(* Logix 5000 project; controller CIP vendor 1 type 14 code 106 rev 20.12; software revision 20.06; part 2 of 13 *)
(* tags used below, declared in another part *)
   Bit : BOOL[128];
   Counter : COUNTER[10];
   IN_N7_100_199 : INT[100];
   Integer : DINT[150];
   Integer_1 : ALIAS FOR Integer[1];
   Level_Bits : BOOL[32];
   One_Shot : BOOL[128];
   OpCode_Pin : DINT[5];
   OpCode_Word : DINT[5,97];
   Panelview : INT[40];
   PV_Security : Security_Main_HMI;
   Recipe : RECIPE[41];

        [24].Setpoint[26] := 9.0, [24].Setpoint[27] := 10.0, [24].Setpoint[28] := 50.0, [24].Setpoint[29] := 3.0, [24].Setpoint[30] := 17.0, [24].Setpoint[31] := 300.0, [24].Setpoint[32] := 2.0, [24].Setpoint[33] := 2.0, [24].Setpoint[34] := 900.0, [24].Setpoint[37] := 70.0, [24].Setpoint[38] := 100.0, [24].Setpoint[39] := 110.0, [24].Setpoint[40] := 30.0, [24].Setpoint[41] := 60.0, [24].Setpoint[42] := 60.0, [24].Setpoint[43] := 3000.0, [24].Setpoint[44] := 300.0, [24].Setpoint[45] := 185.0, [24].Setpoint[46] := 10.0, [24].Setpoint[47] := 25.0, [24].Setpoint[48] := 150.0, [24].Setpoint[49] := 125.0, [24].Setpoint[50] := 100.0, [24].Setpoint[51] := 80.0, [24].Setpoint[52] := 100.0, [24].Setpoint[53] := 50.0, [24].Setpoint[54] := 85.0, [24].Setpoint[55] := 40.0, [24].Setpoint[56] := 60.0, [24].Setpoint[57] := 90.0, [24].Setpoint[58] := 4.0, [24].Setpoint[61] := 10.0, [24].Setpoint[62] := 1.0, [24].Setpoint[65] := 100.0, [24].Setpoint[66] := 15.0, [24].Setpoint[67] := 50.0, [24].Setpoint[68] := 5.0, [24].Setpoint[69] := 100.0, [24].Setpoint[70] := 15.0, [24].Setpoint[71] := 100.0, [24].Setpoint[72] := 15.0, [24].Setpoint[73] := 120.0, [24].Setpoint[74] := 20.0, [24].Setpoint[75] := 120.0, [24].Setpoint[76] := 20.0, [24].Setpoint[77] := 100.0, [24].Setpoint[78] := 15.0, [24].Setpoint[79] := 100.0, [24].Setpoint[80] := 15.0, [24].Setpoint[81] := 45.0, [24].Setpoint[82] := 30.0, [24].Setpoint[83] := 5.0, [24].Setpoint[85] := 5.0, [24].Setpoint[86] := 9.0, [24].Setpoint[92] := 75.0, [24].Setpoint[93] := 90.0, [24].Setpoint[94] := 5.0, [24].Setpoint[95] := 110.0, [24].Setpoint[96] := 10.0, [24].Name := 'RECIPE #24',
        [25].Setpoint[1] := 55.0, [25].Setpoint[2] := 65.0, [25].Setpoint[3] := 60.0, [25].Setpoint[4] := 45.0, [25].Setpoint[5] := 65.0, [25].Setpoint[6] := 25.0, [25].Setpoint[7] := 53.0, [25].Setpoint[8] := 63.0, [25].Setpoint[9] := 57.0, [25].Setpoint[10] := 43.0, [25].Setpoint[11] := 63.0, [25].Setpoint[12] := 22.0, [25].Setpoint[13] := 85.0, [25].Setpoint[14] := 900.0, [25].Setpoint[15] := 300.0, [25].Setpoint[16] := 300.0, [25].Setpoint[17] := 15.0, [25].Setpoint[18] := 14.0, [25].Setpoint[19] := 15.0, [25].Setpoint[20] := 45.0, [25].Setpoint[21] := 5.0, [25].Setpoint[22] := 15.0, [25].Setpoint[23] := 300.0, [25].Setpoint[24] := 2.0, [25].Setpoint[25] := 10.0, [25].Setpoint[26] := 9.0, [25].Setpoint[27] := 10.0, [25].Setpoint[28] := 50.0, [25].Setpoint[29] := 3.0, [25].Setpoint[30] := 17.0, [25].Setpoint[31] := 300.0, [25].Setpoint[32] := 2.0, [25].Setpoint[33] := 2.0, [25].Setpoint[34] := 900.0, [25].Setpoint[37] := 70.0, [25].Setpoint[38] := 100.0, [25].Setpoint[39] := 110.0, [25].Setpoint[40] := 30.0, [25].Setpoint[41] := 60.0, [25].Setpoint[42] := 60.0, [25].Setpoint[43] := 3000.0, [25].Setpoint[44] := 300.0, [25].Setpoint[45] := 185.0, [25].Setpoint[46] := 10.0, [25].Setpoint[47] := 25.0, [25].Setpoint[48] := 150.0, [25].Setpoint[49] := 125.0, [25].Setpoint[50] := 100.0, [25].Setpoint[51] := 80.0, [25].Setpoint[52] := 100.0, [25].Setpoint[53] := 50.0, [25].Setpoint[54] := 85.0, [25].Setpoint[55] := 40.0, [25].Setpoint[56] := 60.0, [25].Setpoint[57] := 90.0, [25].Setpoint[58] := 4.0, [25].Setpoint[61] := 10.0, [25].Setpoint[62] := 1.0, [25].Setpoint[65] := 100.0, [25].Setpoint[66] := 15.0,
        [25].Setpoint[67] := 50.0, [25].Setpoint[68] := 5.0, [25].Setpoint[69] := 100.0, [25].Setpoint[70] := 15.0, [25].Setpoint[71] := 100.0, [25].Setpoint[72] := 15.0, [25].Setpoint[73] := 120.0, [25].Setpoint[74] := 20.0, [25].Setpoint[75] := 120.0, [25].Setpoint[76] := 20.0, [25].Setpoint[77] := 100.0, [25].Setpoint[78] := 15.0, [25].Setpoint[79] := 100.0, [25].Setpoint[80] := 15.0, [25].Setpoint[81] := 45.0, [25].Setpoint[82] := 30.0, [25].Setpoint[83] := 5.0, [25].Setpoint[85] := 5.0, [25].Setpoint[86] := 9.0, [25].Setpoint[92] := 75.0, [25].Setpoint[93] := 90.0, [25].Setpoint[94] := 5.0, [25].Setpoint[95] := 110.0, [25].Setpoint[96] := 10.0, [25].Name := 'RECIPE #25', [26].Setpoint[1] := 55.0, [26].Setpoint[2] := 65.0, [26].Setpoint[3] := 60.0, [26].Setpoint[4] := 45.0, [26].Setpoint[5] := 65.0, [26].Setpoint[6] := 25.0, [26].Setpoint[7] := 53.0, [26].Setpoint[8] := 63.0, [26].Setpoint[9] := 57.0, [26].Setpoint[10] := 43.0, [26].Setpoint[11] := 63.0, [26].Setpoint[12] := 22.0, [26].Setpoint[13] := 85.0, [26].Setpoint[14] := 900.0, [26].Setpoint[15] := 300.0, [26].Setpoint[16] := 300.0, [26].Setpoint[17] := 15.0, [26].Setpoint[18] := 14.0, [26].Setpoint[19] := 15.0, [26].Setpoint[20] := 45.0, [26].Setpoint[21] := 5.0, [26].Setpoint[22] := 15.0, [26].Setpoint[23] := 300.0, [26].Setpoint[24] := 2.0, [26].Setpoint[25] := 10.0, [26].Setpoint[26] := 9.0, [26].Setpoint[27] := 10.0, [26].Setpoint[28] := 50.0, [26].Setpoint[29] := 3.0, [26].Setpoint[30] := 17.0, [26].Setpoint[31] := 300.0, [26].Setpoint[32] := 2.0, [26].Setpoint[33] := 2.0, [26].Setpoint[34] := 900.0, [26].Setpoint[37] := 70.0,
        [26].Setpoint[38] := 100.0, [26].Setpoint[39] := 110.0, [26].Setpoint[40] := 30.0, [26].Setpoint[41] := 60.0, [26].Setpoint[42] := 60.0, [26].Setpoint[43] := 3000.0, [26].Setpoint[44] := 300.0, [26].Setpoint[45] := 185.0, [26].Setpoint[46] := 10.0, [26].Setpoint[47] := 25.0, [26].Setpoint[48] := 150.0, [26].Setpoint[49] := 125.0, [26].Setpoint[50] := 100.0, [26].Setpoint[51] := 80.0, [26].Setpoint[52] := 100.0, [26].Setpoint[53] := 50.0, [26].Setpoint[54] := 85.0, [26].Setpoint[55] := 40.0, [26].Setpoint[56] := 60.0, [26].Setpoint[57] := 90.0, [26].Setpoint[58] := 4.0, [26].Setpoint[61] := 10.0, [26].Setpoint[62] := 1.0, [26].Setpoint[65] := 100.0, [26].Setpoint[66] := 15.0, [26].Setpoint[67] := 50.0, [26].Setpoint[68] := 5.0, [26].Setpoint[69] := 100.0, [26].Setpoint[70] := 15.0, [26].Setpoint[71] := 100.0, [26].Setpoint[72] := 15.0, [26].Setpoint[73] := 120.0, [26].Setpoint[74] := 20.0, [26].Setpoint[75] := 120.0, [26].Setpoint[76] := 20.0, [26].Setpoint[77] := 100.0, [26].Setpoint[78] := 15.0, [26].Setpoint[79] := 100.0, [26].Setpoint[80] := 15.0, [26].Setpoint[81] := 45.0, [26].Setpoint[82] := 30.0, [26].Setpoint[83] := 5.0, [26].Setpoint[85] := 5.0, [26].Setpoint[86] := 9.0, [26].Setpoint[92] := 75.0, [26].Setpoint[93] := 90.0, [26].Setpoint[94] := 5.0, [26].Setpoint[95] := 110.0, [26].Setpoint[96] := 10.0, [26].Name := 'RECIPE #26', [27].Setpoint[1] := 55.0, [27].Setpoint[2] := 65.0, [27].Setpoint[3] := 60.0, [27].Setpoint[4] := 45.0, [27].Setpoint[5] := 65.0, [27].Setpoint[6] := 25.0, [27].Setpoint[7] := 53.0, [27].Setpoint[8] := 63.0, [27].Setpoint[9] := 57.0, [27].Setpoint[10] := 43.0,
        [27].Setpoint[11] := 63.0, [27].Setpoint[12] := 22.0, [27].Setpoint[13] := 85.0, [27].Setpoint[14] := 900.0, [27].Setpoint[15] := 300.0, [27].Setpoint[16] := 300.0, [27].Setpoint[17] := 15.0, [27].Setpoint[18] := 14.0, [27].Setpoint[19] := 15.0, [27].Setpoint[20] := 45.0, [27].Setpoint[21] := 5.0, [27].Setpoint[22] := 15.0, [27].Setpoint[23] := 300.0, [27].Setpoint[24] := 2.0, [27].Setpoint[25] := 10.0, [27].Setpoint[26] := 9.0, [27].Setpoint[27] := 10.0, [27].Setpoint[28] := 50.0, [27].Setpoint[29] := 3.0, [27].Setpoint[30] := 17.0, [27].Setpoint[31] := 300.0, [27].Setpoint[32] := 2.0, [27].Setpoint[33] := 2.0, [27].Setpoint[34] := 900.0, [27].Setpoint[37] := 70.0, [27].Setpoint[38] := 100.0, [27].Setpoint[39] := 110.0, [27].Setpoint[40] := 30.0, [27].Setpoint[41] := 60.0, [27].Setpoint[42] := 60.0, [27].Setpoint[43] := 3000.0, [27].Setpoint[44] := 300.0, [27].Setpoint[45] := 185.0, [27].Setpoint[46] := 10.0, [27].Setpoint[47] := 25.0, [27].Setpoint[48] := 150.0, [27].Setpoint[49] := 125.0, [27].Setpoint[50] := 100.0, [27].Setpoint[51] := 80.0, [27].Setpoint[52] := 100.0, [27].Setpoint[53] := 50.0, [27].Setpoint[54] := 85.0, [27].Setpoint[55] := 40.0, [27].Setpoint[56] := 60.0, [27].Setpoint[57] := 90.0, [27].Setpoint[58] := 4.0, [27].Setpoint[61] := 10.0, [27].Setpoint[62] := 1.0, [27].Setpoint[65] := 100.0, [27].Setpoint[66] := 15.0, [27].Setpoint[67] := 50.0, [27].Setpoint[68] := 5.0, [27].Setpoint[69] := 100.0, [27].Setpoint[70] := 15.0, [27].Setpoint[71] := 100.0, [27].Setpoint[72] := 15.0, [27].Setpoint[73] := 120.0, [27].Setpoint[74] := 20.0, [27].Setpoint[75] := 120.0, [27].Setpoint[76] := 20.0,
        [27].Setpoint[77] := 100.0, [27].Setpoint[78] := 15.0, [27].Setpoint[79] := 100.0, [27].Setpoint[80] := 15.0, [27].Setpoint[81] := 45.0, [27].Setpoint[82] := 30.0, [27].Setpoint[83] := 5.0, [27].Setpoint[85] := 5.0, [27].Setpoint[86] := 9.0, [27].Setpoint[92] := 75.0, [27].Setpoint[93] := 90.0, [27].Setpoint[94] := 5.0, [27].Setpoint[95] := 110.0, [27].Setpoint[96] := 10.0, [27].Name := 'RECIPE #27', [28].Setpoint[1] := 55.0, [28].Setpoint[2] := 65.0, [28].Setpoint[3] := 60.0, [28].Setpoint[4] := 45.0, [28].Setpoint[5] := 65.0, [28].Setpoint[6] := 25.0, [28].Setpoint[7] := 53.0, [28].Setpoint[8] := 63.0, [28].Setpoint[9] := 57.0, [28].Setpoint[10] := 43.0, [28].Setpoint[11] := 63.0, [28].Setpoint[12] := 22.0, [28].Setpoint[13] := 85.0, [28].Setpoint[14] := 900.0, [28].Setpoint[15] := 300.0, [28].Setpoint[16] := 300.0, [28].Setpoint[17] := 15.0, [28].Setpoint[18] := 14.0, [28].Setpoint[19] := 15.0, [28].Setpoint[20] := 45.0, [28].Setpoint[21] := 5.0, [28].Setpoint[22] := 15.0, [28].Setpoint[23] := 300.0, [28].Setpoint[24] := 2.0, [28].Setpoint[25] := 10.0, [28].Setpoint[26] := 9.0, [28].Setpoint[27] := 10.0, [28].Setpoint[28] := 50.0, [28].Setpoint[29] := 3.0, [28].Setpoint[30] := 17.0, [28].Setpoint[31] := 300.0, [28].Setpoint[32] := 2.0, [28].Setpoint[33] := 2.0, [28].Setpoint[34] := 900.0, [28].Setpoint[37] := 70.0, [28].Setpoint[38] := 100.0, [28].Setpoint[39] := 110.0, [28].Setpoint[40] := 30.0, [28].Setpoint[41] := 60.0, [28].Setpoint[42] := 60.0, [28].Setpoint[43] := 3000.0, [28].Setpoint[44] := 300.0, [28].Setpoint[45] := 185.0, [28].Setpoint[46] := 10.0, [28].Setpoint[47] := 25.0,
        [28].Setpoint[48] := 150.0, [28].Setpoint[49] := 125.0, [28].Setpoint[50] := 100.0, [28].Setpoint[51] := 80.0, [28].Setpoint[52] := 100.0, [28].Setpoint[53] := 50.0, [28].Setpoint[54] := 85.0, [28].Setpoint[55] := 40.0, [28].Setpoint[56] := 60.0, [28].Setpoint[57] := 90.0, [28].Setpoint[58] := 4.0, [28].Setpoint[61] := 10.0, [28].Setpoint[62] := 1.0, [28].Setpoint[65] := 100.0, [28].Setpoint[66] := 15.0, [28].Setpoint[67] := 50.0, [28].Setpoint[68] := 5.0, [28].Setpoint[69] := 100.0, [28].Setpoint[70] := 15.0, [28].Setpoint[71] := 100.0, [28].Setpoint[72] := 15.0, [28].Setpoint[73] := 120.0, [28].Setpoint[74] := 20.0, [28].Setpoint[75] := 120.0, [28].Setpoint[76] := 20.0, [28].Setpoint[77] := 100.0, [28].Setpoint[78] := 15.0, [28].Setpoint[79] := 100.0, [28].Setpoint[80] := 15.0, [28].Setpoint[81] := 45.0, [28].Setpoint[82] := 30.0, [28].Setpoint[83] := 5.0, [28].Setpoint[85] := 5.0, [28].Setpoint[86] := 9.0, [28].Setpoint[92] := 75.0, [28].Setpoint[93] := 90.0, [28].Setpoint[94] := 5.0, [28].Setpoint[95] := 110.0, [28].Setpoint[96] := 10.0, [28].Name := 'RECIPE #28', [29].Setpoint[1] := 55.0, [29].Setpoint[2] := 65.0, [29].Setpoint[3] := 60.0, [29].Setpoint[4] := 45.0, [29].Setpoint[5] := 65.0, [29].Setpoint[6] := 25.0, [29].Setpoint[7] := 53.0, [29].Setpoint[8] := 63.0, [29].Setpoint[9] := 57.0, [29].Setpoint[10] := 43.0, [29].Setpoint[11] := 63.0, [29].Setpoint[12] := 22.0, [29].Setpoint[13] := 85.0, [29].Setpoint[14] := 900.0, [29].Setpoint[15] := 300.0, [29].Setpoint[16] := 300.0, [29].Setpoint[17] := 15.0, [29].Setpoint[18] := 14.0, [29].Setpoint[19] := 15.0, [29].Setpoint[20] := 45.0,
        [29].Setpoint[21] := 5.0, [29].Setpoint[22] := 15.0, [29].Setpoint[23] := 300.0, [29].Setpoint[24] := 2.0, [29].Setpoint[25] := 10.0, [29].Setpoint[26] := 9.0, [29].Setpoint[27] := 10.0, [29].Setpoint[28] := 50.0, [29].Setpoint[29] := 3.0, [29].Setpoint[30] := 17.0, [29].Setpoint[31] := 300.0, [29].Setpoint[32] := 2.0, [29].Setpoint[33] := 2.0, [29].Setpoint[34] := 900.0, [29].Setpoint[37] := 70.0, [29].Setpoint[38] := 100.0, [29].Setpoint[39] := 110.0, [29].Setpoint[40] := 30.0, [29].Setpoint[41] := 60.0, [29].Setpoint[42] := 60.0, [29].Setpoint[43] := 3000.0, [29].Setpoint[44] := 300.0, [29].Setpoint[45] := 185.0, [29].Setpoint[46] := 10.0, [29].Setpoint[47] := 25.0, [29].Setpoint[48] := 150.0, [29].Setpoint[49] := 125.0, [29].Setpoint[50] := 100.0, [29].Setpoint[51] := 80.0, [29].Setpoint[52] := 100.0, [29].Setpoint[53] := 50.0, [29].Setpoint[54] := 85.0, [29].Setpoint[55] := 40.0, [29].Setpoint[56] := 60.0, [29].Setpoint[57] := 90.0, [29].Setpoint[58] := 4.0, [29].Setpoint[61] := 10.0, [29].Setpoint[62] := 1.0, [29].Setpoint[65] := 100.0, [29].Setpoint[66] := 15.0, [29].Setpoint[67] := 50.0, [29].Setpoint[68] := 5.0, [29].Setpoint[69] := 100.0, [29].Setpoint[70] := 15.0, [29].Setpoint[71] := 100.0, [29].Setpoint[72] := 15.0, [29].Setpoint[73] := 120.0, [29].Setpoint[74] := 20.0, [29].Setpoint[75] := 120.0, [29].Setpoint[76] := 20.0, [29].Setpoint[77] := 100.0, [29].Setpoint[78] := 15.0, [29].Setpoint[79] := 100.0, [29].Setpoint[80] := 15.0, [29].Setpoint[81] := 45.0, [29].Setpoint[82] := 30.0, [29].Setpoint[83] := 5.0, [29].Setpoint[85] := 5.0, [29].Setpoint[86] := 9.0, [29].Setpoint[92] := 75.0,
        [29].Setpoint[93] := 90.0, [29].Setpoint[94] := 5.0, [29].Setpoint[95] := 110.0, [29].Setpoint[96] := 10.0, [29].Name := 'RECIPE #29', [30].Setpoint[1] := 55.0, [30].Setpoint[2] := 65.0, [30].Setpoint[3] := 60.0, [30].Setpoint[4] := 45.0, [30].Setpoint[5] := 65.0, [30].Setpoint[6] := 25.0, [30].Setpoint[7] := 53.0, [30].Setpoint[8] := 63.0, [30].Setpoint[9] := 57.0, [30].Setpoint[10] := 43.0, [30].Setpoint[11] := 63.0, [30].Setpoint[12] := 22.0, [30].Setpoint[13] := 85.0, [30].Setpoint[14] := 900.0, [30].Setpoint[15] := 300.0, [30].Setpoint[16] := 300.0, [30].Setpoint[17] := 15.0, [30].Setpoint[18] := 14.0, [30].Setpoint[19] := 15.0, [30].Setpoint[20] := 45.0, [30].Setpoint[21] := 5.0, [30].Setpoint[22] := 15.0, [30].Setpoint[23] := 300.0, [30].Setpoint[24] := 2.0, [30].Setpoint[25] := 10.0, [30].Setpoint[26] := 9.0, [30].Setpoint[27] := 10.0, [30].Setpoint[28] := 50.0, [30].Setpoint[29] := 3.0, [30].Setpoint[30] := 17.0, [30].Setpoint[31] := 300.0, [30].Setpoint[32] := 2.0, [30].Setpoint[33] := 2.0, [30].Setpoint[34] := 900.0, [30].Setpoint[37] := 70.0, [30].Setpoint[38] := 100.0, [30].Setpoint[39] := 110.0, [30].Setpoint[40] := 30.0, [30].Setpoint[41] := 60.0, [30].Setpoint[42] := 60.0, [30].Setpoint[43] := 3000.0, [30].Setpoint[44] := 300.0, [30].Setpoint[45] := 185.0, [30].Setpoint[46] := 10.0, [30].Setpoint[47] := 25.0, [30].Setpoint[48] := 150.0, [30].Setpoint[49] := 125.0, [30].Setpoint[50] := 100.0, [30].Setpoint[51] := 80.0, [30].Setpoint[52] := 100.0, [30].Setpoint[53] := 50.0, [30].Setpoint[54] := 85.0, [30].Setpoint[55] := 40.0, [30].Setpoint[56] := 60.0, [30].Setpoint[57] := 90.0,
        [30].Setpoint[58] := 4.0, [30].Setpoint[61] := 10.0, [30].Setpoint[62] := 1.0, [30].Setpoint[65] := 100.0, [30].Setpoint[66] := 15.0, [30].Setpoint[67] := 50.0, [30].Setpoint[68] := 5.0, [30].Setpoint[69] := 100.0, [30].Setpoint[70] := 15.0, [30].Setpoint[71] := 100.0, [30].Setpoint[72] := 15.0, [30].Setpoint[73] := 120.0, [30].Setpoint[74] := 20.0, [30].Setpoint[75] := 120.0, [30].Setpoint[76] := 20.0, [30].Setpoint[77] := 100.0, [30].Setpoint[78] := 15.0, [30].Setpoint[79] := 100.0, [30].Setpoint[80] := 15.0, [30].Setpoint[81] := 45.0, [30].Setpoint[82] := 30.0, [30].Setpoint[83] := 5.0, [30].Setpoint[85] := 5.0, [30].Setpoint[86] := 9.0, [30].Setpoint[92] := 75.0, [30].Setpoint[93] := 90.0, [30].Setpoint[94] := 5.0, [30].Setpoint[95] := 110.0, [30].Setpoint[96] := 10.0, [30].Name := 'RECIPE #30', [31].Setpoint[1] := 55.0, [31].Setpoint[2] := 65.0, [31].Setpoint[3] := 60.0, [31].Setpoint[4] := 45.0, [31].Setpoint[5] := 65.0, [31].Setpoint[6] := 25.0, [31].Setpoint[7] := 53.0, [31].Setpoint[8] := 63.0, [31].Setpoint[9] := 57.0, [31].Setpoint[10] := 43.0, [31].Setpoint[11] := 63.0, [31].Setpoint[12] := 22.0, [31].Setpoint[13] := 85.0, [31].Setpoint[14] := 900.0, [31].Setpoint[15] := 300.0, [31].Setpoint[16] := 300.0, [31].Setpoint[17] := 15.0, [31].Setpoint[18] := 14.0, [31].Setpoint[19] := 15.0, [31].Setpoint[20] := 45.0, [31].Setpoint[21] := 5.0, [31].Setpoint[22] := 15.0, [31].Setpoint[23] := 300.0, [31].Setpoint[24] := 2.0, [31].Setpoint[25] := 10.0, [31].Setpoint[26] := 9.0, [31].Setpoint[27] := 10.0, [31].Setpoint[28] := 50.0, [31].Setpoint[29] := 3.0, [31].Setpoint[30] := 17.0,
        [31].Setpoint[31] := 300.0, [31].Setpoint[32] := 2.0, [31].Setpoint[33] := 2.0, [31].Setpoint[34] := 900.0, [31].Setpoint[37] := 70.0, [31].Setpoint[38] := 100.0, [31].Setpoint[39] := 110.0, [31].Setpoint[40] := 30.0, [31].Setpoint[41] := 60.0, [31].Setpoint[42] := 60.0, [31].Setpoint[43] := 3000.0, [31].Setpoint[44] := 300.0, [31].Setpoint[45] := 185.0, [31].Setpoint[46] := 10.0, [31].Setpoint[47] := 25.0, [31].Setpoint[48] := 150.0, [31].Setpoint[49] := 125.0, [31].Setpoint[50] := 100.0, [31].Setpoint[51] := 80.0, [31].Setpoint[52] := 100.0, [31].Setpoint[53] := 50.0, [31].Setpoint[54] := 85.0, [31].Setpoint[55] := 40.0, [31].Setpoint[56] := 60.0, [31].Setpoint[57] := 90.0, [31].Setpoint[58] := 4.0, [31].Setpoint[61] := 10.0, [31].Setpoint[62] := 1.0, [31].Setpoint[65] := 100.0, [31].Setpoint[66] := 15.0, [31].Setpoint[67] := 50.0, [31].Setpoint[68] := 5.0, [31].Setpoint[69] := 100.0, [31].Setpoint[70] := 15.0, [31].Setpoint[71] := 100.0, [31].Setpoint[72] := 15.0, [31].Setpoint[73] := 120.0, [31].Setpoint[74] := 20.0, [31].Setpoint[75] := 120.0, [31].Setpoint[76] := 20.0, [31].Setpoint[77] := 100.0, [31].Setpoint[78] := 15.0, [31].Setpoint[79] := 100.0, [31].Setpoint[80] := 15.0, [31].Setpoint[81] := 45.0, [31].Setpoint[82] := 30.0, [31].Setpoint[83] := 5.0, [31].Setpoint[85] := 5.0, [31].Setpoint[86] := 9.0, [31].Setpoint[92] := 75.0, [31].Setpoint[93] := 90.0, [31].Setpoint[94] := 5.0, [31].Setpoint[95] := 110.0, [31].Setpoint[96] := 10.0, [31].Name := 'RECIPE #31', [32].Setpoint[1] := 55.0, [32].Setpoint[2] := 65.0, [32].Setpoint[3] := 60.0, [32].Setpoint[4] := 45.0, [32].Setpoint[5] := 65.0,
        [32].Setpoint[6] := 25.0, [32].Setpoint[7] := 53.0, [32].Setpoint[8] := 63.0, [32].Setpoint[9] := 57.0, [32].Setpoint[10] := 43.0, [32].Setpoint[11] := 63.0, [32].Setpoint[12] := 22.0, [32].Setpoint[13] := 85.0, [32].Setpoint[14] := 900.0, [32].Setpoint[15] := 300.0, [32].Setpoint[16] := 300.0, [32].Setpoint[17] := 15.0, [32].Setpoint[18] := 14.0, [32].Setpoint[19] := 15.0, [32].Setpoint[20] := 45.0, [32].Setpoint[21] := 5.0, [32].Setpoint[22] := 15.0, [32].Setpoint[23] := 300.0, [32].Setpoint[24] := 2.0, [32].Setpoint[25] := 10.0, [32].Setpoint[26] := 9.0, [32].Setpoint[27] := 10.0, [32].Setpoint[28] := 50.0, [32].Setpoint[29] := 3.0, [32].Setpoint[30] := 17.0, [32].Setpoint[31] := 300.0, [32].Setpoint[32] := 2.0, [32].Setpoint[33] := 2.0, [32].Setpoint[34] := 900.0, [32].Setpoint[37] := 70.0, [32].Setpoint[38] := 100.0, [32].Setpoint[39] := 110.0, [32].Setpoint[40] := 30.0, [32].Setpoint[41] := 60.0, [32].Setpoint[42] := 60.0, [32].Setpoint[43] := 3000.0, [32].Setpoint[44] := 300.0, [32].Setpoint[45] := 185.0, [32].Setpoint[46] := 10.0, [32].Setpoint[47] := 25.0, [32].Setpoint[48] := 150.0, [32].Setpoint[49] := 125.0, [32].Setpoint[50] := 100.0, [32].Setpoint[51] := 80.0, [32].Setpoint[52] := 100.0, [32].Setpoint[53] := 50.0, [32].Setpoint[54] := 85.0, [32].Setpoint[55] := 40.0, [32].Setpoint[56] := 60.0, [32].Setpoint[57] := 90.0, [32].Setpoint[58] := 4.0, [32].Setpoint[61] := 10.0, [32].Setpoint[62] := 1.0, [32].Setpoint[65] := 100.0, [32].Setpoint[66] := 15.0, [32].Setpoint[67] := 50.0, [32].Setpoint[68] := 5.0, [32].Setpoint[69] := 100.0, [32].Setpoint[70] := 15.0, [32].Setpoint[71] := 100.0,
        [32].Setpoint[72] := 15.0, [32].Setpoint[73] := 120.0, [32].Setpoint[74] := 20.0, [32].Setpoint[75] := 120.0, [32].Setpoint[76] := 20.0, [32].Setpoint[77] := 100.0, [32].Setpoint[78] := 15.0, [32].Setpoint[79] := 100.0, [32].Setpoint[80] := 15.0, [32].Setpoint[81] := 45.0, [32].Setpoint[82] := 30.0, [32].Setpoint[83] := 5.0, [32].Setpoint[85] := 5.0, [32].Setpoint[86] := 9.0, [32].Setpoint[92] := 75.0, [32].Setpoint[93] := 90.0, [32].Setpoint[94] := 5.0, [32].Setpoint[95] := 110.0, [32].Setpoint[96] := 10.0, [32].Name := 'RECIPE #32', [33].Setpoint[1] := 55.0, [33].Setpoint[2] := 65.0, [33].Setpoint[3] := 60.0, [33].Setpoint[4] := 45.0, [33].Setpoint[5] := 65.0, [33].Setpoint[6] := 25.0, [33].Setpoint[7] := 53.0, [33].Setpoint[8] := 63.0, [33].Setpoint[9] := 57.0, [33].Setpoint[10] := 43.0, [33].Setpoint[11] := 63.0, [33].Setpoint[12] := 22.0, [33].Setpoint[13] := 85.0, [33].Setpoint[14] := 900.0, [33].Setpoint[15] := 300.0, [33].Setpoint[16] := 300.0, [33].Setpoint[17] := 15.0, [33].Setpoint[18] := 14.0, [33].Setpoint[19] := 15.0, [33].Setpoint[20] := 45.0, [33].Setpoint[21] := 5.0, [33].Setpoint[22] := 15.0, [33].Setpoint[23] := 300.0, [33].Setpoint[24] := 2.0, [33].Setpoint[25] := 10.0, [33].Setpoint[26] := 9.0, [33].Setpoint[27] := 10.0, [33].Setpoint[28] := 50.0, [33].Setpoint[29] := 3.0, [33].Setpoint[30] := 17.0, [33].Setpoint[31] := 300.0, [33].Setpoint[32] := 2.0, [33].Setpoint[33] := 2.0, [33].Setpoint[34] := 900.0, [33].Setpoint[37] := 70.0, [33].Setpoint[38] := 100.0, [33].Setpoint[39] := 110.0, [33].Setpoint[40] := 30.0, [33].Setpoint[41] := 60.0, [33].Setpoint[42] := 60.0,
        [33].Setpoint[43] := 3000.0, [33].Setpoint[44] := 300.0, [33].Setpoint[45] := 185.0, [33].Setpoint[46] := 10.0, [33].Setpoint[47] := 25.0, [33].Setpoint[48] := 150.0, [33].Setpoint[49] := 125.0, [33].Setpoint[50] := 100.0, [33].Setpoint[51] := 80.0, [33].Setpoint[52] := 100.0, [33].Setpoint[53] := 50.0, [33].Setpoint[54] := 85.0, [33].Setpoint[55] := 40.0, [33].Setpoint[56] := 60.0, [33].Setpoint[57] := 90.0, [33].Setpoint[58] := 4.0, [33].Setpoint[61] := 10.0, [33].Setpoint[62] := 1.0, [33].Setpoint[65] := 100.0, [33].Setpoint[66] := 15.0, [33].Setpoint[67] := 50.0, [33].Setpoint[68] := 5.0, [33].Setpoint[69] := 100.0, [33].Setpoint[70] := 15.0, [33].Setpoint[71] := 100.0, [33].Setpoint[72] := 15.0, [33].Setpoint[73] := 120.0, [33].Setpoint[74] := 20.0, [33].Setpoint[75] := 120.0, [33].Setpoint[76] := 20.0, [33].Setpoint[77] := 100.0, [33].Setpoint[78] := 15.0, [33].Setpoint[79] := 100.0, [33].Setpoint[80] := 15.0, [33].Setpoint[81] := 45.0, [33].Setpoint[82] := 30.0, [33].Setpoint[83] := 5.0, [33].Setpoint[85] := 5.0, [33].Setpoint[86] := 9.0, [33].Setpoint[92] := 75.0, [33].Setpoint[93] := 90.0, [33].Setpoint[94] := 5.0, [33].Setpoint[95] := 110.0, [33].Setpoint[96] := 10.0, [33].Name := 'RECIPE #33', [34].Setpoint[1] := 55.0, [34].Setpoint[2] := 65.0, [34].Setpoint[3] := 60.0, [34].Setpoint[4] := 45.0, [34].Setpoint[5] := 65.0, [34].Setpoint[6] := 25.0, [34].Setpoint[7] := 53.0, [34].Setpoint[8] := 63.0, [34].Setpoint[9] := 57.0, [34].Setpoint[10] := 43.0, [34].Setpoint[11] := 63.0, [34].Setpoint[12] := 22.0, [34].Setpoint[13] := 85.0, [34].Setpoint[14] := 900.0, [34].Setpoint[15] := 300.0,
        [34].Setpoint[16] := 300.0, [34].Setpoint[17] := 15.0, [34].Setpoint[18] := 14.0, [34].Setpoint[19] := 15.0, [34].Setpoint[20] := 45.0, [34].Setpoint[21] := 5.0, [34].Setpoint[22] := 15.0, [34].Setpoint[23] := 300.0, [34].Setpoint[24] := 2.0, [34].Setpoint[25] := 10.0, [34].Setpoint[26] := 9.0, [34].Setpoint[27] := 10.0, [34].Setpoint[28] := 50.0, [34].Setpoint[29] := 3.0, [34].Setpoint[30] := 17.0, [34].Setpoint[31] := 300.0, [34].Setpoint[32] := 2.0, [34].Setpoint[33] := 2.0, [34].Setpoint[34] := 900.0, [34].Setpoint[37] := 70.0, [34].Setpoint[38] := 100.0, [34].Setpoint[39] := 110.0, [34].Setpoint[40] := 30.0, [34].Setpoint[41] := 60.0, [34].Setpoint[42] := 60.0, [34].Setpoint[43] := 3000.0, [34].Setpoint[44] := 300.0, [34].Setpoint[45] := 185.0, [34].Setpoint[46] := 10.0, [34].Setpoint[47] := 25.0, [34].Setpoint[48] := 150.0, [34].Setpoint[49] := 125.0, [34].Setpoint[50] := 100.0, [34].Setpoint[51] := 80.0, [34].Setpoint[52] := 100.0, [34].Setpoint[53] := 50.0, [34].Setpoint[54] := 85.0, [34].Setpoint[55] := 40.0, [34].Setpoint[56] := 60.0, [34].Setpoint[57] := 90.0, [34].Setpoint[58] := 4.0, [34].Setpoint[61] := 10.0, [34].Setpoint[62] := 1.0, [34].Setpoint[65] := 100.0, [34].Setpoint[66] := 15.0, [34].Setpoint[67] := 50.0, [34].Setpoint[68] := 5.0, [34].Setpoint[69] := 100.0, [34].Setpoint[70] := 15.0, [34].Setpoint[71] := 100.0, [34].Setpoint[72] := 15.0, [34].Setpoint[73] := 120.0, [34].Setpoint[74] := 20.0, [34].Setpoint[75] := 120.0, [34].Setpoint[76] := 20.0, [34].Setpoint[77] := 100.0, [34].Setpoint[78] := 15.0, [34].Setpoint[79] := 100.0, [34].Setpoint[80] := 15.0, [34].Setpoint[81] := 45.0,
        [34].Setpoint[82] := 30.0, [34].Setpoint[83] := 5.0, [34].Setpoint[85] := 5.0, [34].Setpoint[86] := 9.0, [34].Setpoint[92] := 75.0, [34].Setpoint[93] := 90.0, [34].Setpoint[94] := 5.0, [34].Setpoint[95] := 110.0, [34].Setpoint[96] := 10.0, [34].Name := 'RECIPE #34', [35].Setpoint[1] := 55.0, [35].Setpoint[2] := 65.0, [35].Setpoint[3] := 60.0, [35].Setpoint[4] := 45.0, [35].Setpoint[5] := 65.0, [35].Setpoint[6] := 25.0, [35].Setpoint[7] := 53.0, [35].Setpoint[8] := 63.0, [35].Setpoint[9] := 57.0, [35].Setpoint[10] := 43.0, [35].Setpoint[11] := 63.0, [35].Setpoint[12] := 22.0, [35].Setpoint[13] := 85.0, [35].Setpoint[14] := 900.0, [35].Setpoint[15] := 300.0, [35].Setpoint[16] := 300.0, [35].Setpoint[17] := 15.0, [35].Setpoint[18] := 14.0, [35].Setpoint[19] := 15.0, [35].Setpoint[20] := 45.0, [35].Setpoint[21] := 5.0, [35].Setpoint[22] := 15.0, [35].Setpoint[23] := 300.0, [35].Setpoint[24] := 2.0, [35].Setpoint[25] := 10.0, [35].Setpoint[26] := 9.0, [35].Setpoint[27] := 10.0, [35].Setpoint[28] := 50.0, [35].Setpoint[29] := 3.0, [35].Setpoint[30] := 17.0, [35].Setpoint[31] := 300.0, [35].Setpoint[32] := 2.0, [35].Setpoint[33] := 2.0, [35].Setpoint[34] := 900.0, [35].Setpoint[37] := 70.0, [35].Setpoint[38] := 100.0, [35].Setpoint[39] := 110.0, [35].Setpoint[40] := 30.0, [35].Setpoint[41] := 60.0, [35].Setpoint[42] := 60.0, [35].Setpoint[43] := 3000.0, [35].Setpoint[44] := 300.0, [35].Setpoint[45] := 185.0, [35].Setpoint[46] := 10.0, [35].Setpoint[47] := 25.0, [35].Setpoint[48] := 150.0, [35].Setpoint[49] := 125.0, [35].Setpoint[50] := 100.0, [35].Setpoint[51] := 80.0, [35].Setpoint[52] := 100.0,
        [35].Setpoint[53] := 50.0, [35].Setpoint[54] := 85.0, [35].Setpoint[55] := 40.0, [35].Setpoint[56] := 60.0, [35].Setpoint[57] := 90.0, [35].Setpoint[58] := 4.0, [35].Setpoint[61] := 10.0, [35].Setpoint[62] := 1.0, [35].Setpoint[65] := 100.0, [35].Setpoint[66] := 15.0, [35].Setpoint[67] := 50.0, [35].Setpoint[68] := 5.0, [35].Setpoint[69] := 100.0, [35].Setpoint[70] := 15.0, [35].Setpoint[71] := 100.0, [35].Setpoint[72] := 15.0, [35].Setpoint[73] := 120.0, [35].Setpoint[74] := 20.0, [35].Setpoint[75] := 120.0, [35].Setpoint[76] := 20.0, [35].Setpoint[77] := 100.0, [35].Setpoint[78] := 15.0, [35].Setpoint[79] := 100.0, [35].Setpoint[80] := 15.0, [35].Setpoint[81] := 45.0, [35].Setpoint[82] := 30.0, [35].Setpoint[83] := 5.0, [35].Setpoint[85] := 5.0, [35].Setpoint[86] := 9.0, [35].Setpoint[92] := 75.0, [35].Setpoint[93] := 90.0, [35].Setpoint[94] := 5.0, [35].Setpoint[95] := 110.0, [35].Setpoint[96] := 10.0, [35].Name := 'RECIPE #35', [36].Setpoint[1] := 55.0, [36].Setpoint[2] := 65.0, [36].Setpoint[3] := 60.0, [36].Setpoint[4] := 45.0, [36].Setpoint[5] := 65.0, [36].Setpoint[6] := 25.0, [36].Setpoint[7] := 53.0, [36].Setpoint[8] := 63.0, [36].Setpoint[9] := 57.0, [36].Setpoint[10] := 43.0, [36].Setpoint[11] := 63.0, [36].Setpoint[12] := 22.0, [36].Setpoint[13] := 85.0, [36].Setpoint[14] := 900.0, [36].Setpoint[15] := 300.0, [36].Setpoint[16] := 300.0, [36].Setpoint[17] := 15.0, [36].Setpoint[18] := 14.0, [36].Setpoint[19] := 15.0, [36].Setpoint[20] := 45.0, [36].Setpoint[21] := 5.0, [36].Setpoint[22] := 15.0, [36].Setpoint[23] := 300.0, [36].Setpoint[24] := 2.0, [36].Setpoint[25] := 10.0,
        [36].Setpoint[26] := 9.0, [36].Setpoint[27] := 10.0, [36].Setpoint[28] := 50.0, [36].Setpoint[29] := 3.0, [36].Setpoint[30] := 17.0, [36].Setpoint[31] := 300.0, [36].Setpoint[32] := 2.0, [36].Setpoint[33] := 2.0, [36].Setpoint[34] := 900.0, [36].Setpoint[37] := 70.0, [36].Setpoint[38] := 100.0, [36].Setpoint[39] := 110.0, [36].Setpoint[40] := 30.0, [36].Setpoint[41] := 60.0, [36].Setpoint[42] := 60.0, [36].Setpoint[43] := 3000.0, [36].Setpoint[44] := 300.0, [36].Setpoint[45] := 185.0, [36].Setpoint[46] := 10.0, [36].Setpoint[47] := 25.0, [36].Setpoint[48] := 150.0, [36].Setpoint[49] := 125.0, [36].Setpoint[50] := 100.0, [36].Setpoint[51] := 80.0, [36].Setpoint[52] := 100.0, [36].Setpoint[53] := 50.0, [36].Setpoint[54] := 85.0, [36].Setpoint[55] := 40.0, [36].Setpoint[56] := 60.0, [36].Setpoint[57] := 90.0, [36].Setpoint[58] := 4.0, [36].Setpoint[61] := 10.0, [36].Setpoint[62] := 1.0, [36].Setpoint[65] := 100.0, [36].Setpoint[66] := 15.0, [36].Setpoint[67] := 50.0, [36].Setpoint[68] := 5.0, [36].Setpoint[69] := 100.0, [36].Setpoint[70] := 15.0, [36].Setpoint[71] := 100.0, [36].Setpoint[72] := 15.0, [36].Setpoint[73] := 120.0, [36].Setpoint[74] := 20.0, [36].Setpoint[75] := 120.0, [36].Setpoint[76] := 20.0, [36].Setpoint[77] := 100.0, [36].Setpoint[78] := 15.0, [36].Setpoint[79] := 100.0, [36].Setpoint[80] := 15.0, [36].Setpoint[81] := 45.0, [36].Setpoint[82] := 30.0, [36].Setpoint[83] := 5.0, [36].Setpoint[85] := 5.0, [36].Setpoint[86] := 9.0, [36].Setpoint[92] := 75.0, [36].Setpoint[93] := 90.0, [36].Setpoint[94] := 5.0, [36].Setpoint[95] := 110.0, [36].Setpoint[96] := 10.0, [36].Name := 'RECIPE #36',
        [37].Setpoint[1] := 55.0, [37].Setpoint[2] := 65.0, [37].Setpoint[3] := 60.0, [37].Setpoint[4] := 45.0, [37].Setpoint[5] := 65.0, [37].Setpoint[6] := 25.0, [37].Setpoint[7] := 53.0, [37].Setpoint[8] := 63.0, [37].Setpoint[9] := 57.0, [37].Setpoint[10] := 43.0, [37].Setpoint[11] := 63.0, [37].Setpoint[12] := 22.0, [37].Setpoint[13] := 85.0, [37].Setpoint[14] := 900.0, [37].Setpoint[15] := 300.0, [37].Setpoint[16] := 300.0, [37].Setpoint[17] := 15.0, [37].Setpoint[18] := 14.0, [37].Setpoint[19] := 15.0, [37].Setpoint[20] := 45.0, [37].Setpoint[21] := 5.0, [37].Setpoint[22] := 15.0, [37].Setpoint[23] := 300.0, [37].Setpoint[24] := 2.0, [37].Setpoint[25] := 10.0, [37].Setpoint[26] := 9.0, [37].Setpoint[27] := 10.0, [37].Setpoint[28] := 50.0, [37].Setpoint[29] := 3.0, [37].Setpoint[30] := 17.0, [37].Setpoint[31] := 300.0, [37].Setpoint[32] := 2.0, [37].Setpoint[33] := 2.0, [37].Setpoint[34] := 900.0, [37].Setpoint[37] := 70.0, [37].Setpoint[38] := 100.0, [37].Setpoint[39] := 110.0, [37].Setpoint[40] := 30.0, [37].Setpoint[41] := 60.0, [37].Setpoint[42] := 60.0, [37].Setpoint[43] := 3000.0, [37].Setpoint[44] := 300.0, [37].Setpoint[45] := 185.0, [37].Setpoint[46] := 10.0, [37].Setpoint[47] := 25.0, [37].Setpoint[48] := 150.0, [37].Setpoint[49] := 125.0, [37].Setpoint[50] := 100.0, [37].Setpoint[51] := 80.0, [37].Setpoint[52] := 100.0, [37].Setpoint[53] := 50.0, [37].Setpoint[54] := 85.0, [37].Setpoint[55] := 40.0, [37].Setpoint[56] := 60.0, [37].Setpoint[57] := 90.0, [37].Setpoint[58] := 4.0, [37].Setpoint[61] := 10.0, [37].Setpoint[62] := 1.0, [37].Setpoint[65] := 100.0, [37].Setpoint[66] := 15.0,
        [37].Setpoint[67] := 50.0, [37].Setpoint[68] := 5.0, [37].Setpoint[69] := 100.0, [37].Setpoint[70] := 15.0, [37].Setpoint[71] := 100.0, [37].Setpoint[72] := 15.0, [37].Setpoint[73] := 120.0, [37].Setpoint[74] := 20.0, [37].Setpoint[75] := 120.0, [37].Setpoint[76] := 20.0, [37].Setpoint[77] := 100.0, [37].Setpoint[78] := 15.0, [37].Setpoint[79] := 100.0, [37].Setpoint[80] := 15.0, [37].Setpoint[81] := 45.0, [37].Setpoint[82] := 30.0, [37].Setpoint[83] := 5.0, [37].Setpoint[85] := 5.0, [37].Setpoint[86] := 9.0, [37].Setpoint[92] := 75.0, [37].Setpoint[93] := 90.0, [37].Setpoint[94] := 5.0, [37].Setpoint[95] := 110.0, [37].Setpoint[96] := 10.0, [37].Name := 'RECIPE #37', [38].Setpoint[1] := 55.0, [38].Setpoint[2] := 65.0, [38].Setpoint[3] := 60.0, [38].Setpoint[4] := 45.0, [38].Setpoint[5] := 65.0, [38].Setpoint[6] := 25.0, [38].Setpoint[7] := 53.0, [38].Setpoint[8] := 63.0, [38].Setpoint[9] := 57.0, [38].Setpoint[10] := 43.0, [38].Setpoint[11] := 63.0, [38].Setpoint[12] := 22.0, [38].Setpoint[13] := 85.0, [38].Setpoint[14] := 900.0, [38].Setpoint[15] := 300.0, [38].Setpoint[16] := 300.0, [38].Setpoint[17] := 15.0, [38].Setpoint[18] := 14.0, [38].Setpoint[19] := 15.0, [38].Setpoint[20] := 45.0, [38].Setpoint[21] := 5.0, [38].Setpoint[22] := 15.0, [38].Setpoint[23] := 300.0, [38].Setpoint[24] := 2.0, [38].Setpoint[25] := 10.0, [38].Setpoint[26] := 9.0, [38].Setpoint[27] := 10.0, [38].Setpoint[28] := 50.0, [38].Setpoint[29] := 3.0, [38].Setpoint[30] := 17.0, [38].Setpoint[31] := 300.0, [38].Setpoint[32] := 2.0, [38].Setpoint[33] := 2.0, [38].Setpoint[34] := 900.0, [38].Setpoint[37] := 70.0,
        [38].Setpoint[38] := 100.0, [38].Setpoint[39] := 110.0, [38].Setpoint[40] := 30.0, [38].Setpoint[41] := 60.0, [38].Setpoint[42] := 60.0, [38].Setpoint[43] := 3000.0, [38].Setpoint[44] := 300.0, [38].Setpoint[45] := 185.0, [38].Setpoint[46] := 10.0, [38].Setpoint[47] := 25.0, [38].Setpoint[48] := 150.0, [38].Setpoint[49] := 125.0, [38].Setpoint[50] := 100.0, [38].Setpoint[51] := 80.0, [38].Setpoint[52] := 100.0, [38].Setpoint[53] := 50.0, [38].Setpoint[54] := 85.0, [38].Setpoint[55] := 40.0, [38].Setpoint[56] := 60.0, [38].Setpoint[57] := 90.0, [38].Setpoint[58] := 4.0, [38].Setpoint[61] := 10.0, [38].Setpoint[62] := 1.0, [38].Setpoint[65] := 100.0, [38].Setpoint[66] := 15.0, [38].Setpoint[67] := 50.0, [38].Setpoint[68] := 5.0, [38].Setpoint[69] := 100.0, [38].Setpoint[70] := 15.0, [38].Setpoint[71] := 100.0, [38].Setpoint[72] := 15.0, [38].Setpoint[73] := 120.0, [38].Setpoint[74] := 20.0, [38].Setpoint[75] := 120.0, [38].Setpoint[76] := 20.0, [38].Setpoint[77] := 100.0, [38].Setpoint[78] := 15.0, [38].Setpoint[79] := 100.0, [38].Setpoint[80] := 15.0, [38].Setpoint[81] := 45.0, [38].Setpoint[82] := 30.0, [38].Setpoint[83] := 5.0, [38].Setpoint[85] := 5.0, [38].Setpoint[86] := 9.0, [38].Setpoint[92] := 75.0, [38].Setpoint[93] := 90.0, [38].Setpoint[94] := 5.0, [38].Setpoint[95] := 110.0, [38].Setpoint[96] := 10.0, [38].Name := 'RECIPE #38', [39].Setpoint[1] := 55.0, [39].Setpoint[2] := 65.0, [39].Setpoint[3] := 60.0, [39].Setpoint[4] := 45.0, [39].Setpoint[5] := 65.0, [39].Setpoint[6] := 25.0, [39].Setpoint[7] := 53.0, [39].Setpoint[8] := 63.0, [39].Setpoint[9] := 57.0, [39].Setpoint[10] := 43.0,
        [39].Setpoint[11] := 63.0, [39].Setpoint[12] := 22.0, [39].Setpoint[13] := 85.0, [39].Setpoint[14] := 900.0, [39].Setpoint[15] := 300.0, [39].Setpoint[16] := 300.0, [39].Setpoint[17] := 15.0, [39].Setpoint[18] := 14.0, [39].Setpoint[19] := 15.0, [39].Setpoint[20] := 45.0, [39].Setpoint[21] := 5.0, [39].Setpoint[22] := 15.0, [39].Setpoint[23] := 300.0, [39].Setpoint[24] := 2.0, [39].Setpoint[25] := 10.0, [39].Setpoint[26] := 9.0, [39].Setpoint[27] := 10.0, [39].Setpoint[28] := 50.0, [39].Setpoint[29] := 3.0, [39].Setpoint[30] := 17.0, [39].Setpoint[31] := 300.0, [39].Setpoint[32] := 2.0, [39].Setpoint[33] := 2.0, [39].Setpoint[34] := 900.0, [39].Setpoint[37] := 70.0, [39].Setpoint[38] := 100.0, [39].Setpoint[39] := 110.0, [39].Setpoint[40] := 30.0, [39].Setpoint[41] := 60.0, [39].Setpoint[42] := 60.0, [39].Setpoint[43] := 3000.0, [39].Setpoint[44] := 300.0, [39].Setpoint[45] := 185.0, [39].Setpoint[46] := 10.0, [39].Setpoint[47] := 25.0, [39].Setpoint[48] := 150.0, [39].Setpoint[49] := 125.0, [39].Setpoint[50] := 100.0, [39].Setpoint[51] := 80.0, [39].Setpoint[52] := 100.0, [39].Setpoint[53] := 50.0, [39].Setpoint[54] := 85.0, [39].Setpoint[55] := 40.0, [39].Setpoint[56] := 60.0, [39].Setpoint[57] := 90.0, [39].Setpoint[58] := 4.0, [39].Setpoint[61] := 10.0, [39].Setpoint[62] := 1.0, [39].Setpoint[65] := 100.0, [39].Setpoint[66] := 15.0, [39].Setpoint[67] := 50.0, [39].Setpoint[68] := 5.0, [39].Setpoint[69] := 100.0, [39].Setpoint[70] := 15.0, [39].Setpoint[71] := 100.0, [39].Setpoint[72] := 15.0, [39].Setpoint[73] := 120.0, [39].Setpoint[74] := 20.0, [39].Setpoint[75] := 120.0, [39].Setpoint[76] := 20.0,
        [39].Setpoint[77] := 100.0, [39].Setpoint[78] := 15.0, [39].Setpoint[79] := 100.0, [39].Setpoint[80] := 15.0, [39].Setpoint[81] := 45.0, [39].Setpoint[82] := 30.0, [39].Setpoint[83] := 5.0, [39].Setpoint[85] := 5.0, [39].Setpoint[86] := 9.0, [39].Setpoint[92] := 75.0, [39].Setpoint[93] := 90.0, [39].Setpoint[94] := 5.0, [39].Setpoint[95] := 110.0, [39].Setpoint[96] := 10.0, [39].Name := 'RECIPE #39', [40].Setpoint[1] := 55.0, [40].Setpoint[2] := 65.0, [40].Setpoint[3] := 60.0, [40].Setpoint[4] := 45.0, [40].Setpoint[5] := 65.0, [40].Setpoint[6] := 25.0, [40].Setpoint[7] := 53.0, [40].Setpoint[8] := 63.0, [40].Setpoint[9] := 57.0, [40].Setpoint[10] := 43.0, [40].Setpoint[11] := 63.0, [40].Setpoint[12] := 22.0, [40].Setpoint[13] := 85.0, [40].Setpoint[14] := 900.0, [40].Setpoint[15] := 300.0, [40].Setpoint[16] := 300.0, [40].Setpoint[17] := 15.0, [40].Setpoint[18] := 14.0, [40].Setpoint[19] := 15.0, [40].Setpoint[20] := 45.0, [40].Setpoint[21] := 5.0, [40].Setpoint[22] := 15.0, [40].Setpoint[23] := 300.0, [40].Setpoint[24] := 2.0, [40].Setpoint[25] := 10.0, [40].Setpoint[26] := 9.0, [40].Setpoint[27] := 10.0, [40].Setpoint[28] := 50.0, [40].Setpoint[29] := 3.0, [40].Setpoint[30] := 17.0, [40].Setpoint[31] := 300.0, [40].Setpoint[32] := 2.0, [40].Setpoint[33] := 2.0, [40].Setpoint[34] := 900.0, [40].Setpoint[37] := 25.0, [40].Setpoint[38] := 90.0, [40].Setpoint[39] := 96.0, [40].Setpoint[40] := 60.0, [40].Setpoint[41] := 60.0, [40].Setpoint[42] := 60.0, [40].Setpoint[43] := 3000.0, [40].Setpoint[44] := 300.0, [40].Setpoint[45] := 200.0, [40].Setpoint[46] := 10.0, [40].Setpoint[47] := 25.0,
        [40].Setpoint[48] := 150.0, [40].Setpoint[49] := 125.0, [40].Setpoint[50] := 100.0, [40].Setpoint[51] := 80.0, [40].Setpoint[52] := 100.0, [40].Setpoint[53] := 50.0, [40].Setpoint[54] := 80.0, [40].Setpoint[55] := 40.0, [40].Setpoint[56] := 60.0, [40].Setpoint[57] := 90.0, [40].Setpoint[58] := 4.0, [40].Setpoint[61] := 10.0, [40].Setpoint[62] := 1.0, [40].Setpoint[65] := 100.0, [40].Setpoint[66] := 15.0, [40].Setpoint[67] := 50.0, [40].Setpoint[68] := 5.0, [40].Setpoint[69] := 100.0, [40].Setpoint[70] := 15.0, [40].Setpoint[71] := 100.0, [40].Setpoint[72] := 15.0, [40].Setpoint[73] := 120.0, [40].Setpoint[74] := 20.0, [40].Setpoint[75] := 120.0, [40].Setpoint[76] := 20.0, [40].Setpoint[77] := 100.0, [40].Setpoint[78] := 15.0, [40].Setpoint[79] := 100.0, [40].Setpoint[80] := 15.0, [40].Setpoint[81] := 45.0, [40].Setpoint[82] := 30.0, [40].Setpoint[83] := 5.0, [40].Setpoint[84] := 1.0, [40].Setpoint[85] := 5.0, [40].Setpoint[86] := 9.0, [40].Setpoint[92] := 75.0, [40].Setpoint[93] := 90.0, [40].Setpoint[94] := 5.0, [40].Setpoint[95] := 110.0, [40].Setpoint[96] := 10.0, [40].Name := 'RECIPE #40');
   Recipe_Name : STRING[41] := ([1] := 'TANK WASH W/DIP TUBES CYCLE', [2] := 'TANK WASH W/DIP TUBES CYCLE #2', [3] := 'WASH CHAMBER WASH CYCLE POLY/GLASSWARE', [4] := 'WASH CHAMBER WAS CYCLE PROCESS PARTS', [5] := 'PROCESS HOSES', [6] := 'RECIPE #6', [7] := 'RECIPE #7', [8] := 'RECIPE #8', [9] := 'RECIPE #9', [10] := 'RECIPE #10', [11] := 'RECIPE #11', [12] := 'RECIPE #12', [13] := 'RECIPE #13', [14] := 'RECIPE #14', [15] := 'RECIPE #15', [16] := 'RECIPE #16', [17] := 'RECIPE #17', [18] := 'RECIPE #18', [19] := 'RECIPE #19', [20] := 'RECIPE #20', [21] := 'RECIPE #21', [22] := 'RECIPE #22', [23] := 'RECIPE #23', [24] := 'RECIPE #24', [25] := 'RECIPE #25', [26] := 'RECIPE #26', [27] := 'RECIPE #27', [28] := 'RECIPE #28', [29] := 'RECIPE #29', [30] := 'RECIPE #30', [31] := 'RECIPE #31', [32] := 'RECIPE #32', [33] := 'RECIPE #33', [34] := 'RECIPE #34', [35] := 'RECIPE #35', [36] := 'RECIPE #36', [37] := 'RECIPE #37', [38] := 'RECIPE #38', [39] := 'RECIPE #39', [40] := 'RECIPE #40');
   Recipe_Name_Indx : DINT := 11;
   RotaryONS : DINT;
   SCL_Drain_PH : SCALE := (In := 16546.0, InRawMax := 16383.0, InEUMax := 14.0, Limiting := 1, Out := 14.0, MaxAlarm := 1);
   SCL_Dryer_Duct_Temp : SCALE := (In := 5035.0, InRawMax := 16383.0, InRawMin := 3277.0, InEUMax := 150.0, Out := 20.120556);
   SCL_Dryer_Exhaust_Temp : SCALE := (In := 5028.0, InRawMax := 16383.0, InRawMin := 3277.0, InEUMax := 150.0, Out := 20.04044);
   SCL_Return_Temp : SCALE := (In := 3730.0, InRawMax := 16383.0, InEUMax := 100.0, Out := 22.767504);
   SCL_Rinse_Cond : SCALE := (In := -227.0, InRawMax := 16383.0, InEUMax := 10.0, Limiting := 1, MinAlarm := 1);
   SCL_Solution_Tank_Lvl : SCALE := (In := 3.0, InRawMax := 16383.0, InEUMax := 42.0, Out := 0.007690899);
   SCL_Supply_Flow : SCALE := (In := 344.0, InRawMax := 16383.0, InEUMax := 150.0, Out := 3.1496062);
   SCL_Supply_Flow_CIP_100 : SCALE := (In := -819.0, InRawMax := 16383.0, InEUMax := 30.0, Out := -1.4997253, MinAlarm := 1);
   SCL_Supply_Flow_CIP_200 : SCALE := (In := 3.0, InRawMax := 16383.0, InEUMax := 30.0, Out := 0.0054934993);
   SCL_Supply_Pressure : SCALE := (In := -57.0, InRawMax := 16383.0, InEUMax := 150.0, Out := -0.5218824, MinAlarm := 1);
   SCL_Supply_Temp : SCALE := (In := 3569.0, InRawMax := 16383.0, InEUMax := 100.0, Out := 21.784777);
   SCL_Wash_Chamber_Lvl : SCALE := (In := 3278.0, InRawMax := 16383.0, InRawMin := 3277.0, InEUMax := 12.0, Out := 0.00091561116);
   SCL_Wash_Cond : SCALE := (In := -209.0, InRawMax := 16383.0, InEUMax := 100.0, Limiting := 1, MinAlarm := 1);
   SCLD_Drain_PH : REAL := 14.0;
   SCLD_Dryer_Duct_Temp : REAL := 20.120556;
   SCLD_Dryer_Exhaust_Temp : REAL := 20.051884;
   SCLD_Return_Temp : REAL := 22.761398;
   SCLD_Rinse_Cond : REAL;
   SCLD_Solution_Tank_Lvl : REAL;
   SCLD_Solution_Tank_Lvl_Raw : REAL := 0.007690899;
   SCLD_Supply_Flow : REAL := 3.1587622;
   SCLD_Supply_Flow_CIP : REAL;
   SCLD_Supply_Flow_CIP100 : REAL := -1.4997253;
   SCLD_Supply_Flow_CIP200 : REAL := 0.003662333;
   SCLD_Supply_Pressure : REAL := -0.5218824;
   SCLD_Supply_Temp : REAL := 21.79088;
   SCLD_Wash_Chamber_Lvl : REAL;
   SCLD_Wash_Chamber_Lvl_Raw : REAL;
   SCLD_Wash_Cond : REAL;
   SecurityLevel : DINT;
   SecurityLevel1 : DINT;
   Sequencer : CONTROL[4] := ([0].LEN := 97, [1].LEN := 97, [1].EN := 1, [2].LEN := 6, [3].LEN := 1, [3].POS := 1, [3].DN := 1);
   Solution_Tank_Lvl_Calc : REAL[20] := ([0] := 0.07752426, [1] := 0.14402856, [2] := 0.5431899, [3] := 1.247636, [4] := 2.1940415, [5] := 3.3508313, [6] := 4.8204303, [7] := 6.547088, [8] := 8.440478, [9] := 10.68321, [10] := 13.051815, [11] := 15.73783, [12] := 18.30794, [13] := 21.045364, [14] := 23.834595);
   Solution_Tank_Lvl_Storage : REAL[3];
   SP_Dryer_Min_Temp : REAL;
   SP_Dryer_Temp : REAL;
   SP_Return_Temp : REAL;
   SP_Rinse_Cond : REAL;
   SP_Solution_Tank_Fill_Lvl : REAL := 40.0;
   SP_Solution_Tank_Lvl : REAL := 50.0;
   SP_Supply_Flow : REAL;
   SP_Supply_Temp : REAL;
   SP_Wash_Cond : REAL;
   SP_Wash_Cond_Hold : REAL;
   SP_Wash_Hold_Temp : REAL := 30.0;
   SP_Wash_Temp : REAL := 30.0;
   Time_Date : DINT[20] := ([0] := 2026, [1] := 8, [2] := 24, [3] := 11, [4] := 19, [5] := 3, [6] := 480747, [10] := 2026, [11] := 8, [12] := 24, [13] := 11, [14] := 19, [15] := 3, [16] := 480747);
   Timer : TIMER[99] := ([0].PRE := 2000, [0].ACC := 1234, [0].EN := 1, [0].TT := 1, [1].PRE := 6000, [2].PRE := 2000, [3].PRE := 5000, [4].PRE := 4000, [5].PRE := 20000, [6].PRE := 5000, [7].PRE := 5000, [8].PRE := 6000, [9].PRE := 3600000, [10].PRE := 3000, [11].PRE := 6000, [11].ACC := 6003, [11].EN := 1, [11].DN := 1, [12].PRE := 3000, [12].ACC := 3002, [12].EN := 1, [12].DN := 1, [13].PRE := 1000, [14].PRE := 3000, [15].PRE := 10000, [16].PRE := 20000, [17].PRE := 5000, [18].PRE := 15000, [19].PRE := 5000, [19].ACC := 5000, [19].EN := 1, [19].DN := 1, [20].PRE := 1000, [21].PRE := 5000, [22].PRE := 15000, [23].PRE := 3, [24].PRE := 3, [25].PRE := 3000, [26].PRE := 20000, [27].PRE := 20000, [28].PRE := 20000, [29].PRE := 3, [29].ACC := 3, [30].PRE := 3000, [31].PRE := 1000, [32].PRE := 10000, [33].PRE := 3000, [34].PRE := 1, [35].PRE := 3000, [36].PRE := 20000, [37].PRE := 20000, [38].PRE := 2000, [39].PRE := 5000, [40].PRE := 3000, [40].ACC := 3002, [40].EN := 1, [40].DN := 1, [41].PRE := 10000, [42].PRE := 3000, [42].ACC := 3000,
        [42].EN := 1, [42].TT := 1, [43].PRE := 3000, [43].ACC := 3000, [43].EN := 1, [43].DN := 1, [44].PRE := 10, [45].PRE := 2, [46].PRE := 10, [46].ACC := 9, [47].PRE := 45000, [48].PRE := 45, [49].PRE := 45000, [50].PRE := 5, [51].PRE := 5, [52].PRE := 3, [52].ACC := 3, [53].PRE := 3, [53].ACC := 1, [55].PRE := 75000, [55].ACC := 75001, [55].EN := 1, [55].DN := 1, [56].PRE := 75, [56].ACC := 75, [57].PRE := 300000, [58].PRE := 2000, [59].PRE := 120000, [60].PRE := 100, [60].ACC := 58, [63].PRE := 3000, [63].ACC := 3001, [63].EN := 1, [63].DN := 1, [64].PRE := 2000, [64].ACC := 2001, [64].EN := 1, [64].DN := 1, [65].PRE := 2000, [66].PRE := 300000, [68].PRE := 10000, [68].ACC := 964, [68].EN := 1, [68].TT := 1, [70].PRE := 10000, [70].ACC := 966, [70].EN := 1, [70].TT := 1, [74].PRE := 1000, [74].ACC := 1000, [74].EN := 1, [74].DN := 1, [75].PRE := 1000, [90].PRE := 86400000, [91].PRE := 120000);
   Timer_Chem1_Pump : TIMER[7] := ([0].PRE := 3000, [1].PRE := 30000, [2].PRE := 60000, [3].PRE := 5000, [4].PRE := 15000, [5].PRE := 3000, [5].ACC := 3000);
   Timer_Chem2_Pump : TIMER[7] := ([0].PRE := 3000, [1].PRE := 60000, [2].PRE := 50000, [3].PRE := 30000, [4].PRE := 30000, [5].PRE := 3000, [5].ACC := 3000);
   Utility_Button : DINT[5];
   Utility_Button_ONS : DINT[5];
   Utility_ONS : DINT[5];
   Utility_Out : DINT[5];
   Utility_Timer : TIMER[20] := ([0].PRE := 20000, [1].PRE := 20000, [2].PRE := 20000, [3].PRE := 20000, [4].PRE := 20000, [10].PRE := 20000, [12].PRE := 20000);
   Wash_Chamber_Lvl_Calc : REAL[30] := ([0] := 0.12203876, [1] := 0.20836411, [2] := 0.50576985, [3] := 0.8725683, [4] := 1.3925012, [5] := 2.0347292, [6] := 3.1176043, [7] := 3.8455913, [8] := 5.3291497, [9] := 6.0288644, [10] := 6.7290483, [11] := 8.073697, [12] := 8.739218, [13] := 10.074342, [14] := 11.444196, [15] := 14.314757, [16] := 16.97722, [17] := 20.604128, [18] := 24.562262, [19] := 28.29502, [20] := 32.145573, [21] := 36.29457, [22] := 39.991447, [23] := 44.183628, [24] := 47.83743);
   Wash_Chamber_Lvl_Storage : REAL[3];
   WashChamberDoorGasketCTRL : DINT := 4096;
END_VAR

PROGRAM MainProgram   (* main routine _02_SUB *)

ROUTINE _02_SUB   (* ladder *)
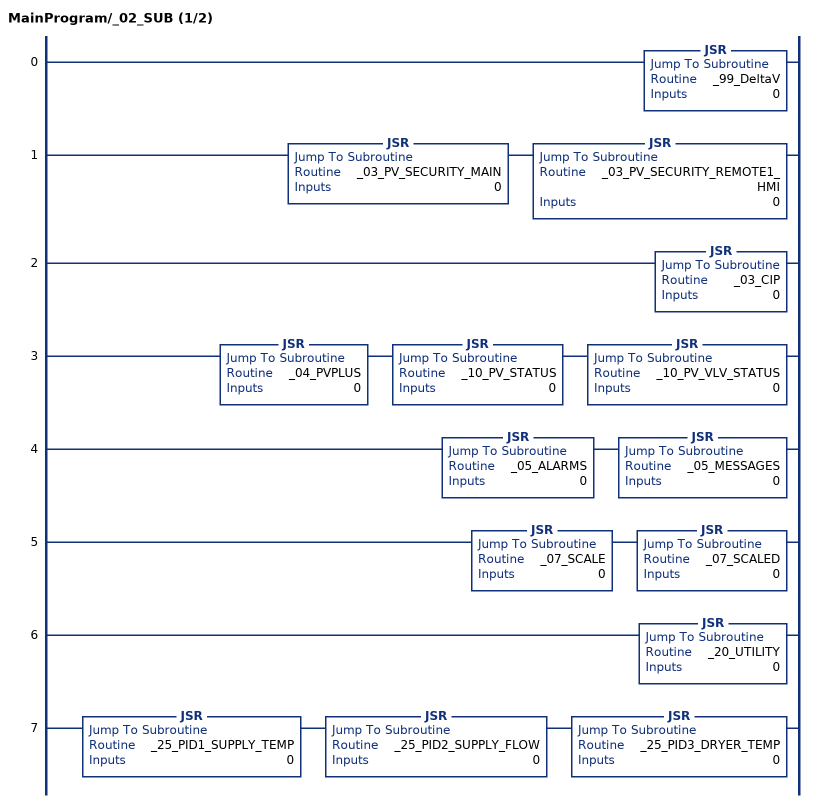
   0: JSR(_99_DeltaV,0);
   1: JSR(_03_PV_SECURITY_MAIN,0)JSR(_03_PV_SECURITY_REMOTE1_HMI,0);
   2: JSR(_03_CIP,0);
   3: JSR(_04_PVPLUS,0)JSR(_10_PV_STATUS,0)JSR(_10_PV_VLV_STATUS,0);
   4: JSR(_05_ALARMS,0)JSR(_05_MESSAGES,0);
   5: JSR(_07_SCALE,0)JSR(_07_SCALED,0);
   6: JSR(_20_UTILITY,0);
   7: JSR(_25_PID1_SUPPLY_TEMP,0)JSR(_25_PID2_SUPPLY_FLOW,0)JSR(_25_PID3_DRYER_TEMP,0);
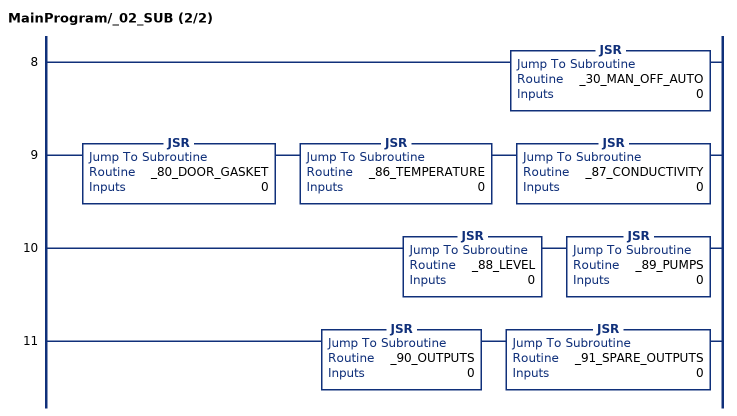
   8: JSR(_30_MAN_OFF_AUTO,0);
   9: JSR(_80_DOOR_GASKET,0)JSR(_86_TEMPERATURE,0)JSR(_87_CONDUCTIVITY,0);
   10: JSR(_88_LEVEL,0)JSR(_89_PUMPS,0);
   11: JSR(_90_OUTPUTS,0)JSR(_91_SPARE_OUTPUTS,0);
END_ROUTINE

ROUTINE _03_CIP   (* ladder *)
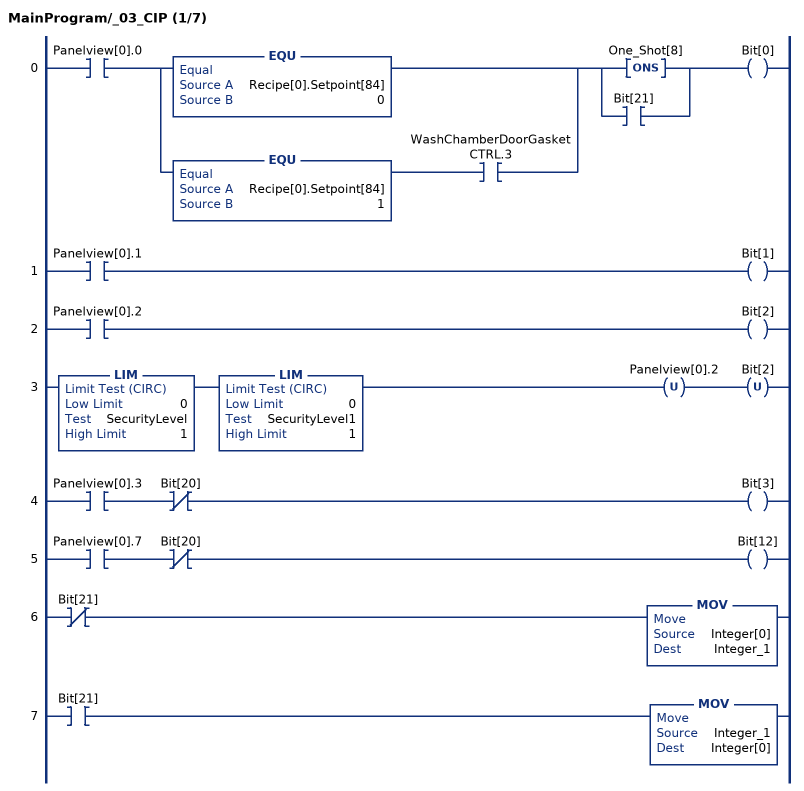
   0: XIC(Panelview[0].0)[EQU(Recipe[0].Setpoint[84],0) ,EQU(Recipe[0].Setpoint[84],1) XIC(WashChamberDoorGasketCTRL.3) ][ONS(One_Shot[8]) ,XIC(Bit[21]) ]OTE(Bit[0]);
   1: XIC(Panelview[0].1)OTE(Bit[1]);
   2: XIC(Panelview[0].2)OTE(Bit[2]);
   3: LIM(0,SecurityLevel,1)LIM(0,SecurityLevel1,1)OTU(Panelview[0].2)OTU(Bit[2]);
   4: XIC(Panelview[0].3)XIO(Bit[20])OTE(Bit[3]);
   5: XIC(Panelview[0].7)XIO(Bit[20])OTE(Bit[12]);
   6: XIO(Bit[21])MOV(Integer[0],Integer_1);
   7: XIC(Bit[21])MOV(Integer_1,Integer[0]);
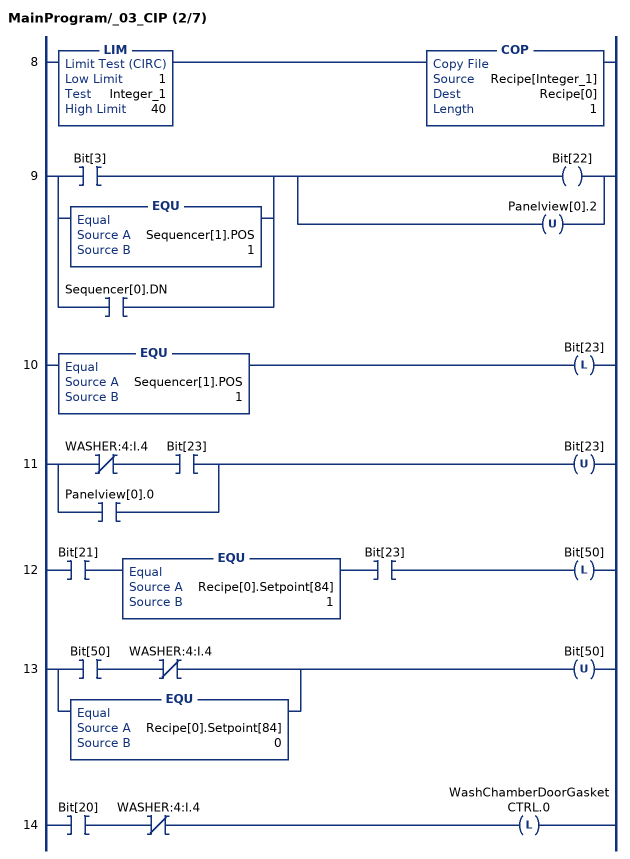
   8: LIM(1,Integer_1,40)COP(Recipe[Integer_1],Recipe[0],1);
   9: [XIC(Bit[3]) ,EQU(Sequencer[1].POS,1) ,XIC(Sequencer[0].DN) ][OTE(Bit[22]) ,OTU(Panelview[0].2) ];
   10: EQU(Sequencer[1].POS,1)OTL(Bit[23]);
   11: [XIO(WASHER:4:I.4) XIC(Bit[23]) ,XIC(Panelview[0].0) ]OTU(Bit[23]);
   12: XIC(Bit[21])EQU(Recipe[0].Setpoint[84],1)XIC(Bit[23])OTL(Bit[50]);
   13: [XIC(Bit[50]) XIO(WASHER:4:I.4) ,EQU(Recipe[0].Setpoint[84],0) ]OTU(Bit[50]);
   14: XIC(Bit[20])XIO(WASHER:4:I.4)OTL(WashChamberDoorGasketCTRL.0);
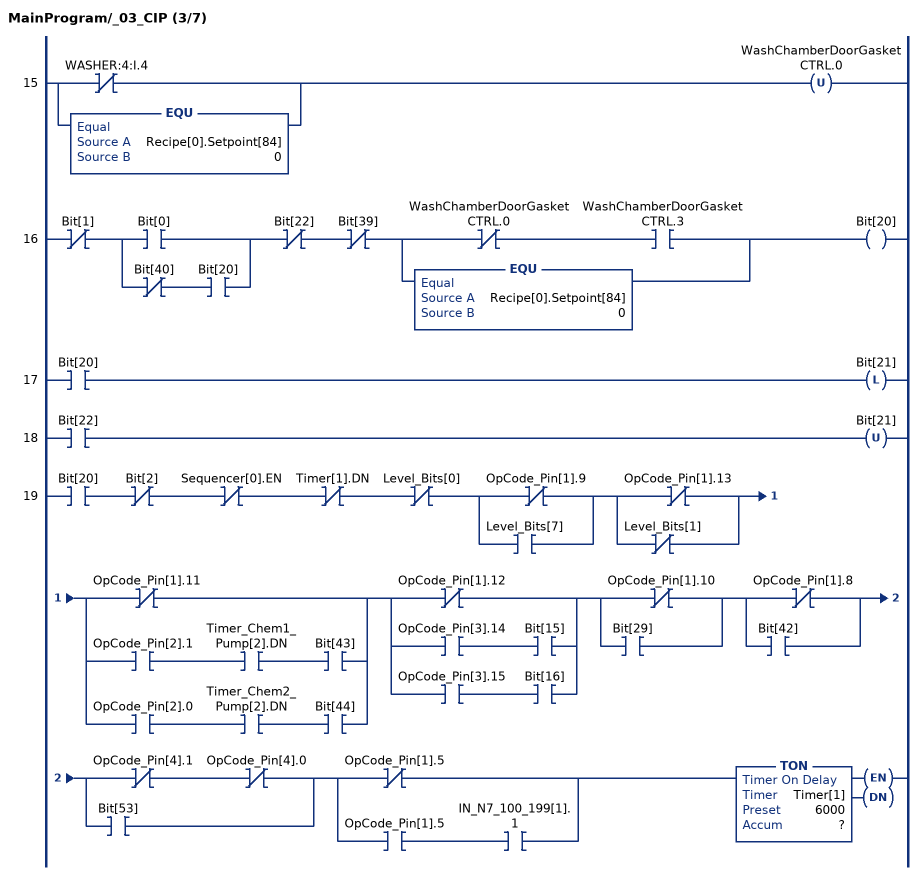
   15: [XIO(WASHER:4:I.4) ,EQU(Recipe[0].Setpoint[84],0) ]OTU(WashChamberDoorGasketCTRL.0);
   16: XIO(Bit[1])[XIC(Bit[0]) ,XIO(Bit[40]) XIC(Bit[20]) ]XIO(Bit[22])XIO(Bit[39])[XIO(WashChamberDoorGasketCTRL.0) XIC(WashChamberDoorGasketCTRL.3) ,EQU(Recipe[0].Setpoint[84],0) ]OTE(Bit[20]);
   17: XIC(Bit[20])OTL(Bit[21]);
   18: XIC(Bit[22])OTU(Bit[21]);
   19: XIC(Bit[20])XIO(Bit[2])XIO(Sequencer[0].EN)XIO(Timer[1].DN)XIO(Level_Bits[0])[XIO(OpCode_Pin[1].9) ,XIC(Level_Bits[7]) ][XIO(OpCode_Pin[1].13) ,XIO(Level_Bits[1]) ][XIO(OpCode_Pin[1].11) ,XIC(OpCode_Pin[2].1) XIC(Timer_Chem1_Pump[2].DN) XIC(Bit[43]) ,XIC(OpCode_Pin[2].0) XIC(Timer_Chem2_Pump[2].DN) XIC(Bit[44]) ][XIO(OpCode_Pin[1].12) ,XIC(OpCode_Pin[3].14) XIC(Bit[15]) ,XIC(OpCode_Pin[3].15) XIC(Bit[16]) ][XIO(OpCode_Pin[1].10) ,XIC(Bit[29]) ][XIO(OpCode_Pin[1].8) ,XIC(Bit[42]) ][XIO(OpCode_Pin[4].1) XIO(OpCode_Pin[4].0) ,XIC(Bit[53]) ][XIO(OpCode_Pin[1].5) ,XIC(OpCode_Pin[1].5) XIC(IN_N7_100_199[1].1) ]TON(Timer[1],?,?);
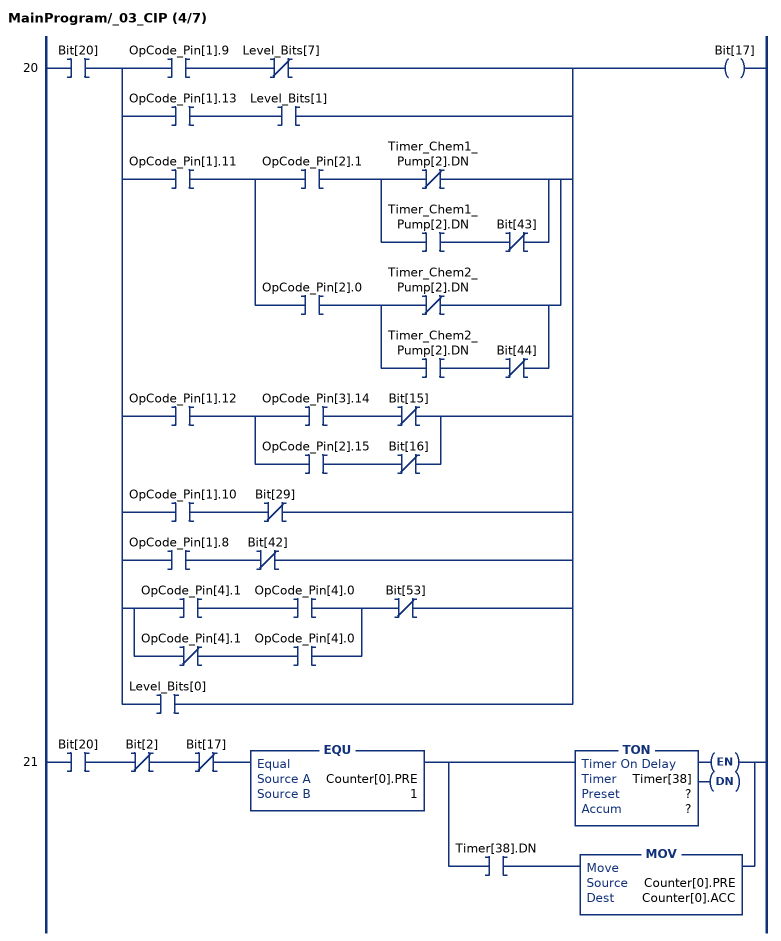
   20: XIC(Bit[20])[XIC(OpCode_Pin[1].9) XIO(Level_Bits[7]) ,XIC(OpCode_Pin[1].13) XIC(Level_Bits[1]) ,XIC(OpCode_Pin[1].11) [XIC(OpCode_Pin[2].1) [XIO(Timer_Chem1_Pump[2].DN) ,XIC(Timer_Chem1_Pump[2].DN) XIO(Bit[43]) ] ,XIC(OpCode_Pin[2].0) [XIO(Timer_Chem2_Pump[2].DN) ,XIC(Timer_Chem2_Pump[2].DN) XIO(Bit[44]) ] ] ,XIC(OpCode_Pin[1].12) [XIC(OpCode_Pin[3].14) XIO(Bit[15]) ,XIC(OpCode_Pin[2].15) XIO(Bit[16]) ] ,XIC(OpCode_Pin[1].10) XIO(Bit[29]) ,XIC(OpCode_Pin[1].8) XIO(Bit[42]) ,[XIC(OpCode_Pin[4].1) XIC(OpCode_Pin[4].0) ,XIO(OpCode_Pin[4].1) XIC(OpCode_Pin[4].0) ] XIO(Bit[53]) ,XIC(Level_Bits[0]) ]OTE(Bit[17]);
   21: XIC(Bit[20])XIO(Bit[2])XIO(Bit[17])EQU(Counter[0].PRE,1)[TON(Timer[38],?,?) ,XIC(Timer[38].DN) MOV(Counter[0].PRE,Counter[0].ACC) ];
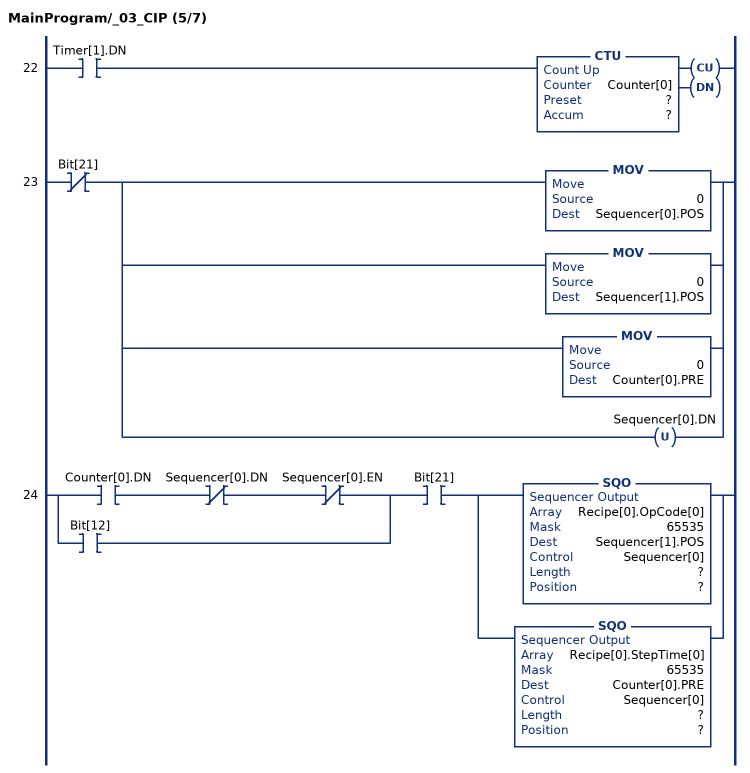
   22: XIC(Timer[1].DN)CTU(Counter[0],?,?);
   23: XIO(Bit[21])[MOV(0,Sequencer[0].POS) ,MOV(0,Sequencer[1].POS) ,MOV(0,Counter[0].PRE) ,OTU(Sequencer[0].DN) ];
   24: [XIC(Counter[0].DN) XIO(Sequencer[0].DN) XIO(Sequencer[0].EN) ,XIC(Bit[12]) ]XIC(Bit[21])[SQO(Recipe[0].OpCode[0],65535,Sequencer[1].POS,Sequencer[0],?,?) ,SQO(Recipe[0].StepTime[0],65535,Counter[0].PRE,Sequencer[0],?,?) ];
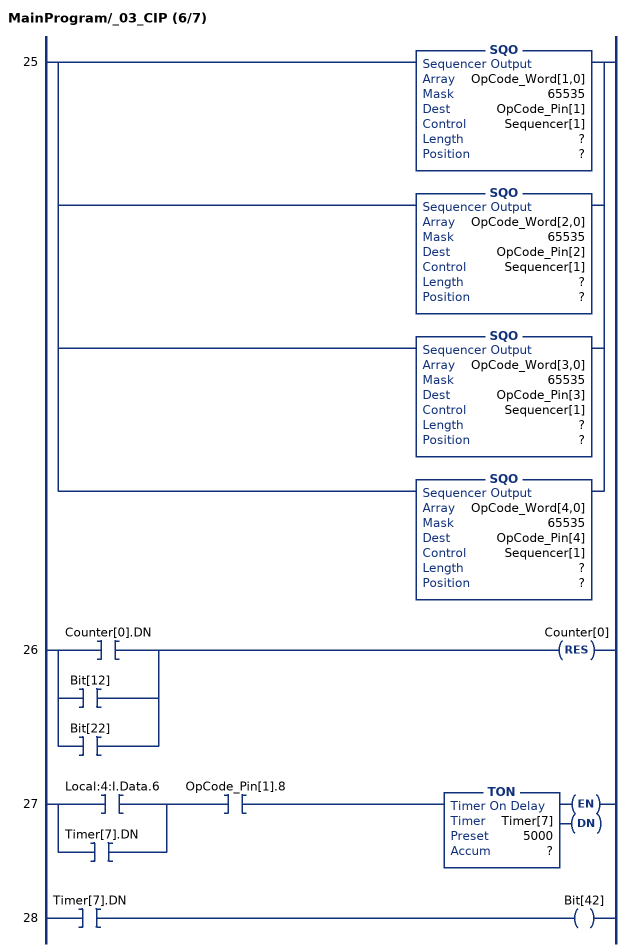
   25: [SQO(OpCode_Word[1,0],65535,OpCode_Pin[1],Sequencer[1],?,?) ,SQO(OpCode_Word[2,0],65535,OpCode_Pin[2],Sequencer[1],?,?) ,SQO(OpCode_Word[3,0],65535,OpCode_Pin[3],Sequencer[1],?,?) ,SQO(OpCode_Word[4,0],65535,OpCode_Pin[4],Sequencer[1],?,?) ];
   26: [XIC(Counter[0].DN) ,XIC(Bit[12]) ,XIC(Bit[22]) ]RES(Counter[0]);
   27: [XIC(Local:4:I.Data.6) ,XIC(Timer[7].DN) ]XIC(OpCode_Pin[1].8)TON(Timer[7],?,?);
   28: XIC(Timer[7].DN)OTE(Bit[42]);
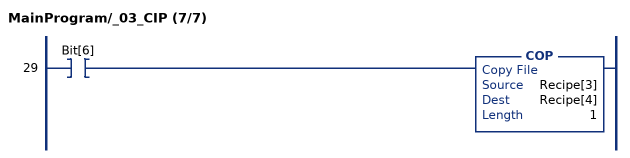
   29: XIC(Bit[6])COP(Recipe[3],Recipe[4],1);
END_ROUTINE

ROUTINE _03_PV_SECURITY_MAIN   (* ladder *)
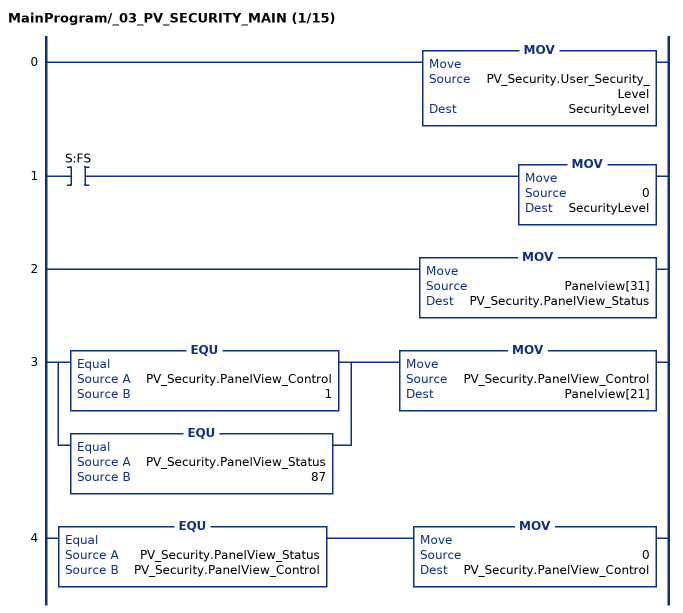
   0: MOV(PV_Security.User_Security_Level,SecurityLevel);
   1: XIC(S:FS)MOV(0,SecurityLevel);
   2: MOV(Panelview[31],PV_Security.PanelView_Status);
   3: [EQU(PV_Security.PanelView_Control,1) ,EQU(PV_Security.PanelView_Status,87) ]MOV(PV_Security.PanelView_Control,Panelview[21]);
   4: EQU(PV_Security.PanelView_Status,PV_Security.PanelView_Control)MOV(0,PV_Security.PanelView_Control);
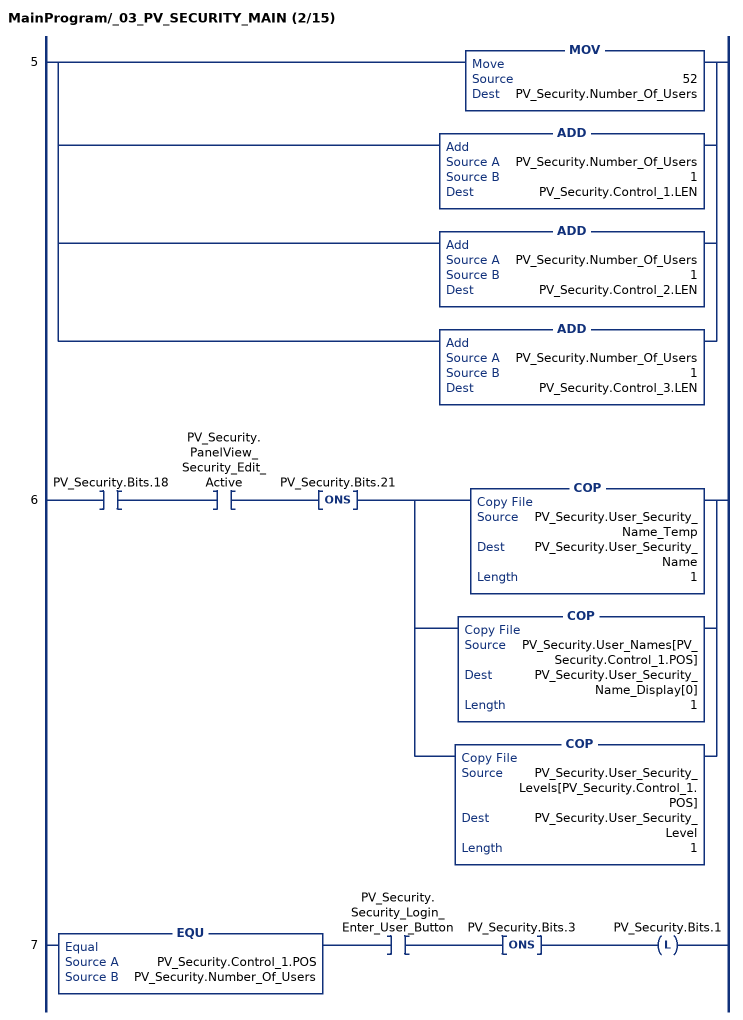
   5: [MOV(52,PV_Security.Number_Of_Users) ,ADD(PV_Security.Number_Of_Users,1,PV_Security.Control_1.LEN) ,ADD(PV_Security.Number_Of_Users,1,PV_Security.Control_2.LEN) ,ADD(PV_Security.Number_Of_Users,1,PV_Security.Control_3.LEN) ];
   6: XIC(PV_Security.Bits.18)XIC(PV_Security.PanelView_Security_Edit_Active)ONS(PV_Security.Bits.21)[COP(PV_Security.User_Security_Name_Temp,PV_Security.User_Security_Name,1) ,COP(PV_Security.User_Names[PV_Security.Control_1.POS],PV_Security.User_Security_Name_Display[0],1) ,COP(PV_Security.User_Security_Levels[PV_Security.Control_1.POS],PV_Security.User_Security_Level,1) ];
   7: EQU(PV_Security.Control_1.POS,PV_Security.Number_Of_Users)XIC(PV_Security.Security_Login_Enter_User_Button)ONS(PV_Security.Bits.3)OTL(PV_Security.Bits.1);
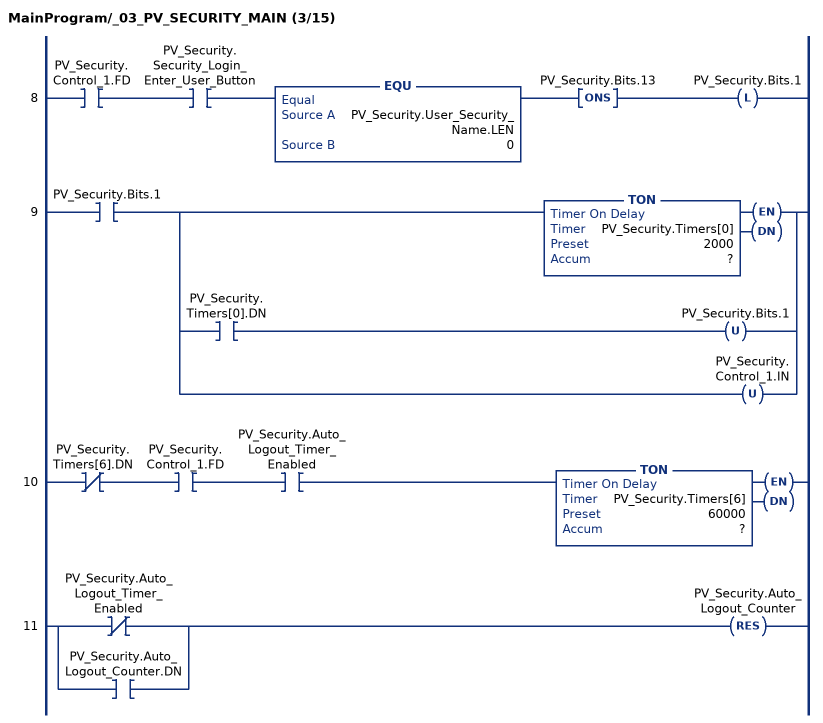
   8: XIC(PV_Security.Control_1.FD)XIC(PV_Security.Security_Login_Enter_User_Button)EQU(PV_Security.User_Security_Name.LEN,0)ONS(PV_Security.Bits.13)OTL(PV_Security.Bits.1);
   9: XIC(PV_Security.Bits.1)[TON(PV_Security.Timers[0],?,?) ,XIC(PV_Security.Timers[0].DN) OTU(PV_Security.Bits.1) ,OTU(PV_Security.Control_1.IN) ];
   10: XIO(PV_Security.Timers[6].DN)XIC(PV_Security.Control_1.FD)XIC(PV_Security.Auto_Logout_Timer_Enabled)TON(PV_Security.Timers[6],?,?);
   11: [XIO(PV_Security.Auto_Logout_Timer_Enabled) ,XIC(PV_Security.Auto_Logout_Counter.DN) ]RES(PV_Security.Auto_Logout_Counter);
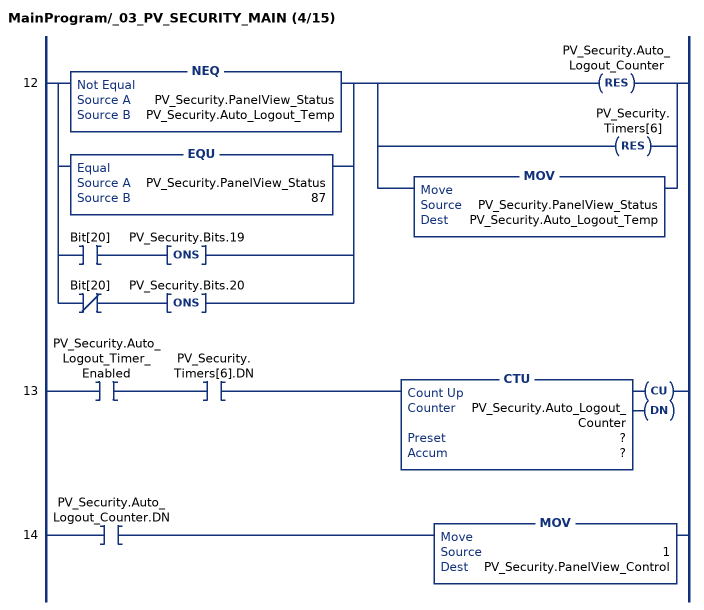
   12: [NEQ(PV_Security.PanelView_Status,PV_Security.Auto_Logout_Temp) ,EQU(PV_Security.PanelView_Status,87) ,XIC(Bit[20]) ONS(PV_Security.Bits.19) ,XIO(Bit[20]) ONS(PV_Security.Bits.20) ][RES(PV_Security.Auto_Logout_Counter) ,RES(PV_Security.Timers[6]) ,MOV(PV_Security.PanelView_Status,PV_Security.Auto_Logout_Temp) ];
   13: XIC(PV_Security.Auto_Logout_Timer_Enabled)XIC(PV_Security.Timers[6].DN)CTU(PV_Security.Auto_Logout_Counter,?,?);
   14: XIC(PV_Security.Auto_Logout_Counter.DN)MOV(1,PV_Security.PanelView_Control);
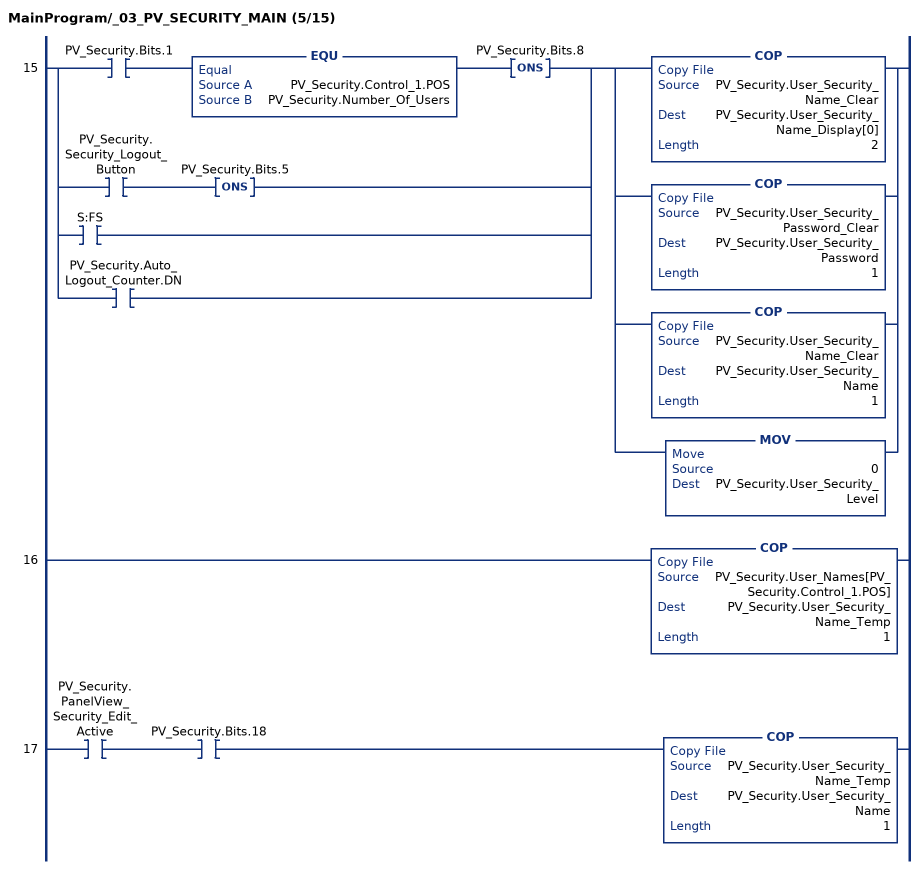
   15: [XIC(PV_Security.Bits.1) EQU(PV_Security.Control_1.POS,PV_Security.Number_Of_Users) ONS(PV_Security.Bits.8) ,XIC(PV_Security.Security_Logout_Button) ONS(PV_Security.Bits.5) ,XIC(S:FS) ,XIC(PV_Security.Auto_Logout_Counter.DN) ][COP(PV_Security.User_Security_Name_Clear,PV_Security.User_Security_Name_Display[0],2) ,COP(PV_Security.User_Security_Password_Clear,PV_Security.User_Security_Password,1) ,COP(PV_Security.User_Security_Name_Clear,PV_Security.User_Security_Name,1) ,MOV(0,PV_Security.User_Security_Level) ];
   16: COP(PV_Security.User_Names[PV_Security.Control_1.POS],PV_Security.User_Security_Name_Temp,1);
   17: XIC(PV_Security.PanelView_Security_Edit_Active)XIC(PV_Security.Bits.18)COP(PV_Security.User_Security_Name_Temp,PV_Security.User_Security_Name,1);
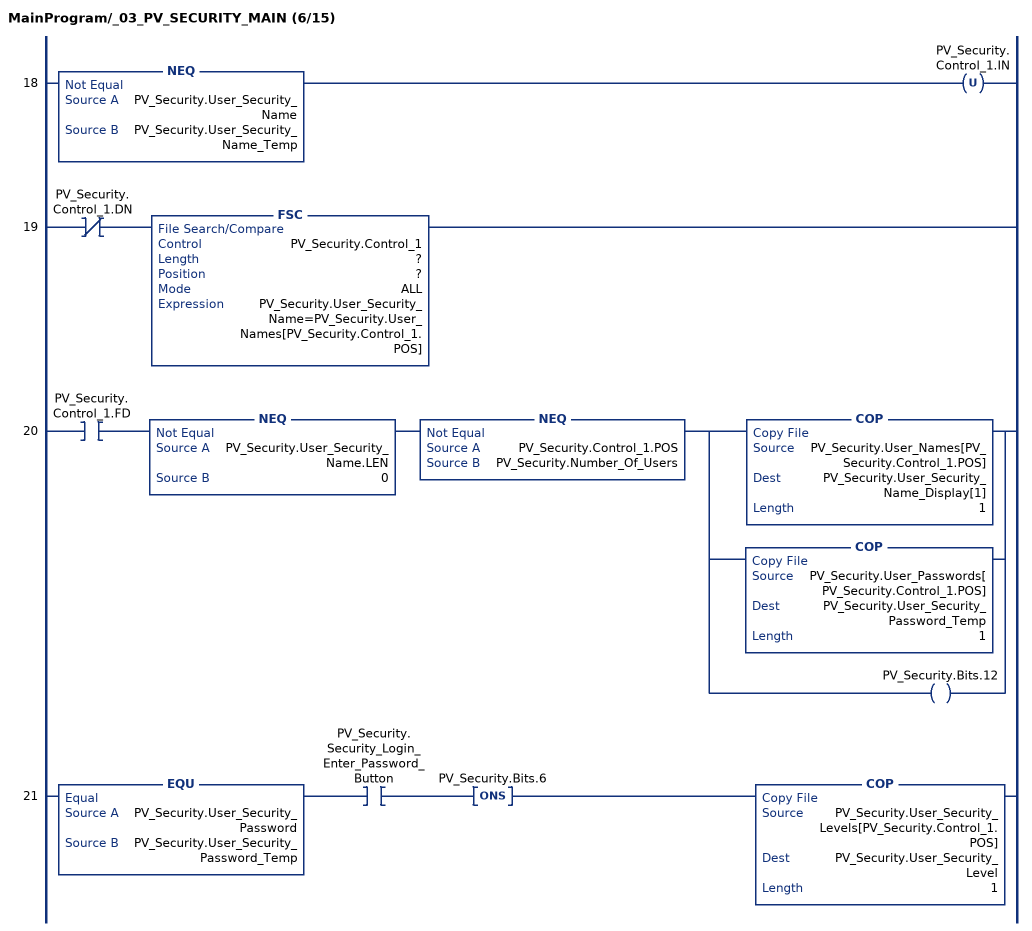
   18: NEQ(PV_Security.User_Security_Name,PV_Security.User_Security_Name_Temp)OTU(PV_Security.Control_1.IN);
   19: XIO(PV_Security.Control_1.DN)FSC(PV_Security.Control_1,?,?,ALL,PV_Security.User_Security_Name=PV_Security.User_Names[PV_Security.Control_1.POS]);
   20: XIC(PV_Security.Control_1.FD)NEQ(PV_Security.User_Security_Name.LEN,0)NEQ(PV_Security.Control_1.POS,PV_Security.Number_Of_Users)[COP(PV_Security.User_Names[PV_Security.Control_1.POS],PV_Security.User_Security_Name_Display[1],1) ,COP(PV_Security.User_Passwords[PV_Security.Control_1.POS],PV_Security.User_Security_Password_Temp,1) ,OTE(PV_Security.Bits.12) ];
   21: EQU(PV_Security.User_Security_Password,PV_Security.User_Security_Password_Temp)XIC(PV_Security.Security_Login_Enter_Password_Button)ONS(PV_Security.Bits.6)COP(PV_Security.User_Security_Levels[PV_Security.Control_1.POS],PV_Security.User_Security_Level,1);
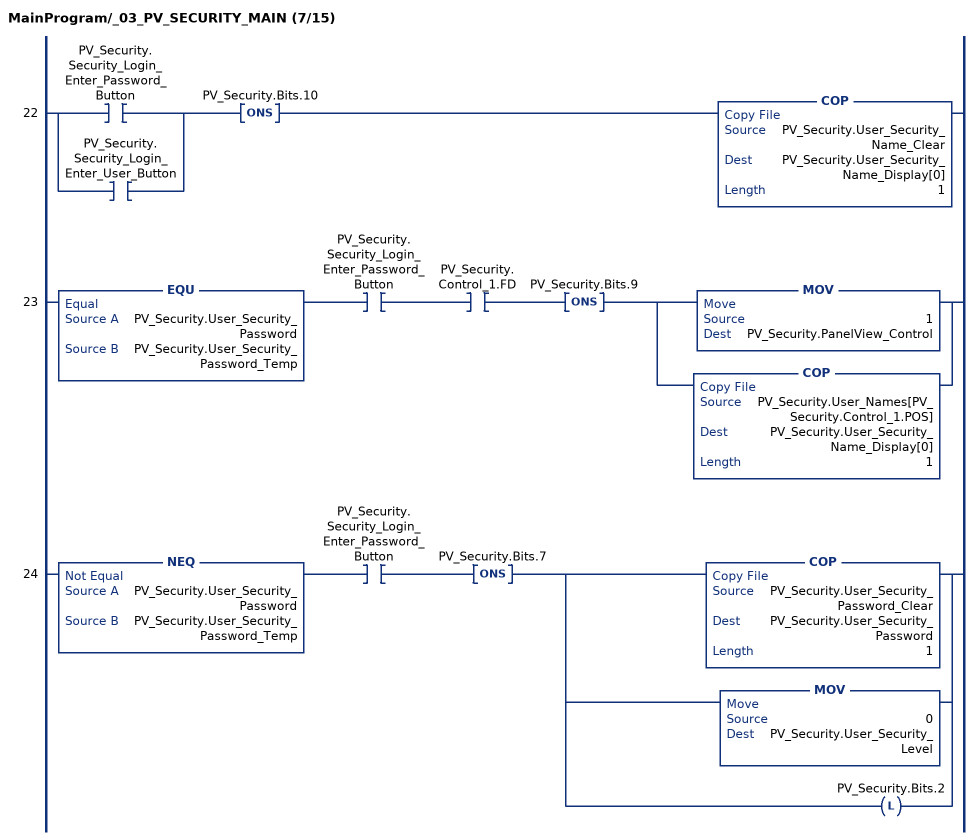
   22: [XIC(PV_Security.Security_Login_Enter_Password_Button) ,XIC(PV_Security.Security_Login_Enter_User_Button) ]ONS(PV_Security.Bits.10)COP(PV_Security.User_Security_Name_Clear,PV_Security.User_Security_Name_Display[0],1);
   23: EQU(PV_Security.User_Security_Password,PV_Security.User_Security_Password_Temp)XIC(PV_Security.Security_Login_Enter_Password_Button)XIC(PV_Security.Control_1.FD)ONS(PV_Security.Bits.9)[MOV(1,PV_Security.PanelView_Control) ,COP(PV_Security.User_Names[PV_Security.Control_1.POS],PV_Security.User_Security_Name_Display[0],1) ];
   24: NEQ(PV_Security.User_Security_Password,PV_Security.User_Security_Password_Temp)XIC(PV_Security.Security_Login_Enter_Password_Button)ONS(PV_Security.Bits.7)[COP(PV_Security.User_Security_Password_Clear,PV_Security.User_Security_Password,1) ,MOV(0,PV_Security.User_Security_Level) ,OTL(PV_Security.Bits.2) ];
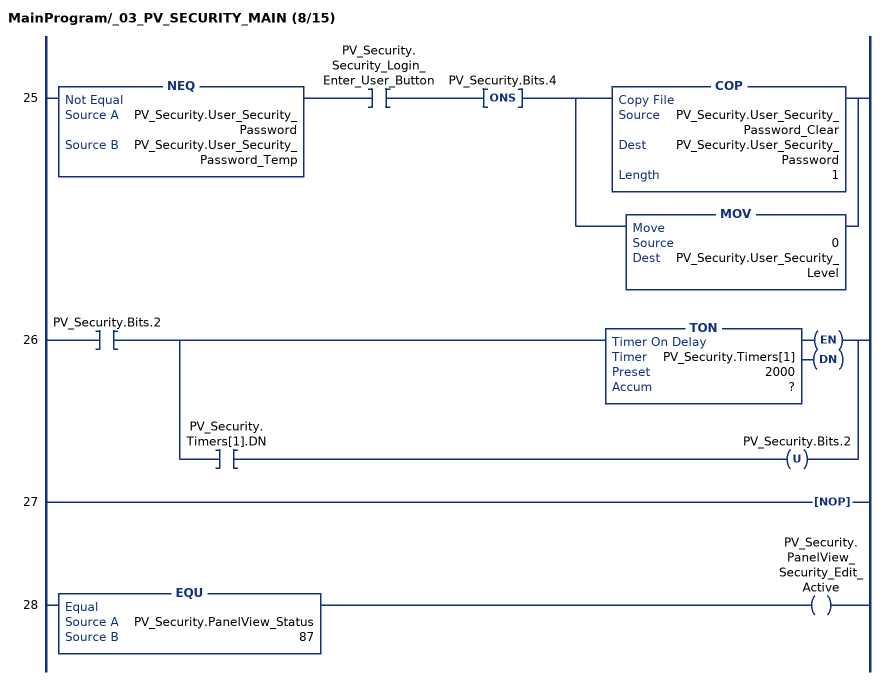
   25: NEQ(PV_Security.User_Security_Password,PV_Security.User_Security_Password_Temp)XIC(PV_Security.Security_Login_Enter_User_Button)ONS(PV_Security.Bits.4)[COP(PV_Security.User_Security_Password_Clear,PV_Security.User_Security_Password,1) ,MOV(0,PV_Security.User_Security_Level) ];
   26: XIC(PV_Security.Bits.2)[TON(PV_Security.Timers[1],?,?) ,XIC(PV_Security.Timers[1].DN) OTU(PV_Security.Bits.2) ];
   27: NOP();
   28: EQU(PV_Security.PanelView_Status,87)OTE(PV_Security.PanelView_Security_Edit_Active);
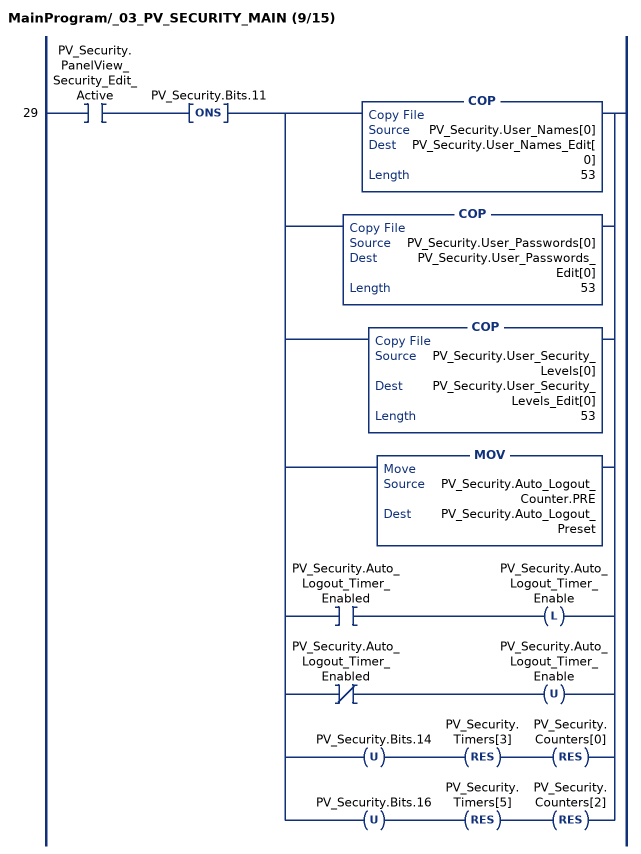
   29: XIC(PV_Security.PanelView_Security_Edit_Active)ONS(PV_Security.Bits.11)[COP(PV_Security.User_Names[0],PV_Security.User_Names_Edit[0],53) ,COP(PV_Security.User_Passwords[0],PV_Security.User_Passwords_Edit[0],53) ,COP(PV_Security.User_Security_Levels[0],PV_Security.User_Security_Levels_Edit[0],53) ,MOV(PV_Security.Auto_Logout_Counter.PRE,PV_Security.Auto_Logout_Preset) ,XIC(PV_Security.Auto_Logout_Timer_Enabled) OTL(PV_Security.Auto_Logout_Timer_Enable) ,XIO(PV_Security.Auto_Logout_Timer_Enabled) OTU(PV_Security.Auto_Logout_Timer_Enable) ,OTU(PV_Security.Bits.14) RES(PV_Security.Timers[3]) RES(PV_Security.Counters[0]) ,OTU(PV_Security.Bits.16) RES(PV_Security.Timers[5]) RES(PV_Security.Counters[2]) ];
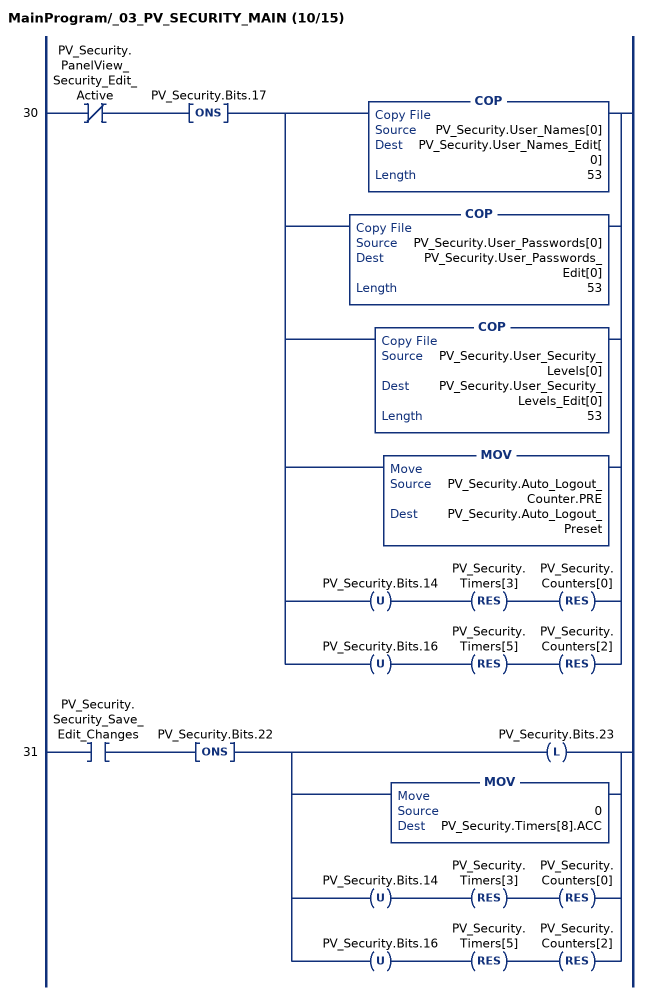
   30: XIO(PV_Security.PanelView_Security_Edit_Active)ONS(PV_Security.Bits.17)[COP(PV_Security.User_Names[0],PV_Security.User_Names_Edit[0],53) ,COP(PV_Security.User_Passwords[0],PV_Security.User_Passwords_Edit[0],53) ,COP(PV_Security.User_Security_Levels[0],PV_Security.User_Security_Levels_Edit[0],53) ,MOV(PV_Security.Auto_Logout_Counter.PRE,PV_Security.Auto_Logout_Preset) ,OTU(PV_Security.Bits.14) RES(PV_Security.Timers[3]) RES(PV_Security.Counters[0]) ,OTU(PV_Security.Bits.16) RES(PV_Security.Timers[5]) RES(PV_Security.Counters[2]) ];
   31: XIC(PV_Security.Security_Save_Edit_Changes)ONS(PV_Security.Bits.22)[OTL(PV_Security.Bits.23) ,MOV(0,PV_Security.Timers[8].ACC) ,OTU(PV_Security.Bits.14) RES(PV_Security.Timers[3]) RES(PV_Security.Counters[0]) ,OTU(PV_Security.Bits.16) RES(PV_Security.Timers[5]) RES(PV_Security.Counters[2]) ];
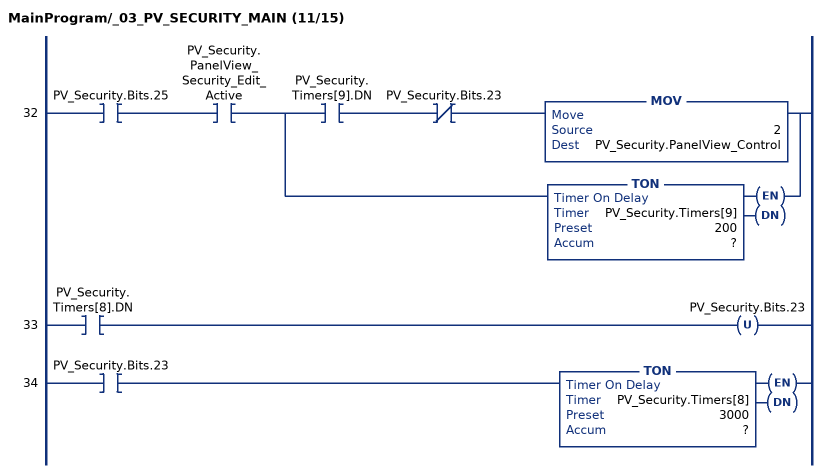
   32: XIC(PV_Security.Bits.25)XIC(PV_Security.PanelView_Security_Edit_Active)[XIC(PV_Security.Timers[9].DN) XIO(PV_Security.Bits.23) MOV(2,PV_Security.PanelView_Control) ,TON(PV_Security.Timers[9],?,?) ];
   33: XIC(PV_Security.Timers[8].DN)OTU(PV_Security.Bits.23);
   34: XIC(PV_Security.Bits.23)TON(PV_Security.Timers[8],?,?);
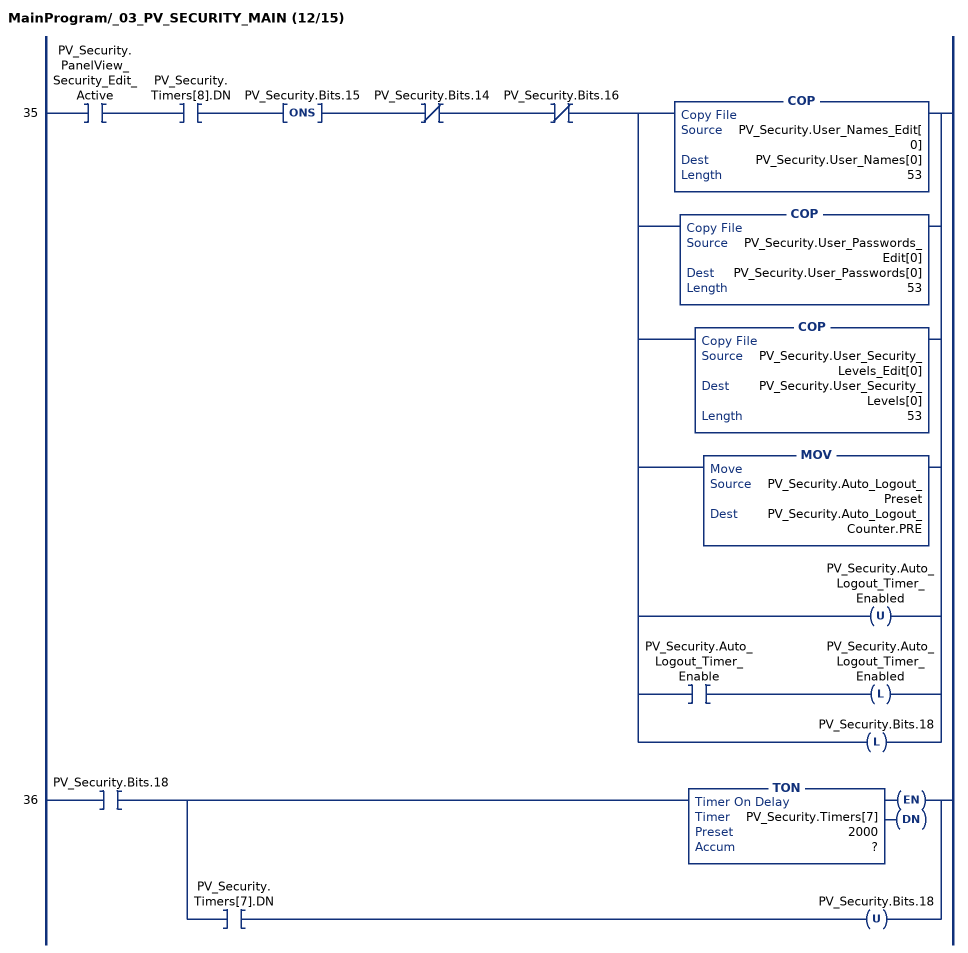
   35: XIC(PV_Security.PanelView_Security_Edit_Active)XIC(PV_Security.Timers[8].DN)ONS(PV_Security.Bits.15)XIO(PV_Security.Bits.14)XIO(PV_Security.Bits.16)[COP(PV_Security.User_Names_Edit[0],PV_Security.User_Names[0],53) ,COP(PV_Security.User_Passwords_Edit[0],PV_Security.User_Passwords[0],53) ,COP(PV_Security.User_Security_Levels_Edit[0],PV_Security.User_Security_Levels[0],53) ,MOV(PV_Security.Auto_Logout_Preset,PV_Security.Auto_Logout_Counter.PRE) ,OTU(PV_Security.Auto_Logout_Timer_Enabled) ,XIC(PV_Security.Auto_Logout_Timer_Enable) OTL(PV_Security.Auto_Logout_Timer_Enabled) ,OTL(PV_Security.Bits.18) ];
   36: XIC(PV_Security.Bits.18)[TON(PV_Security.Timers[7],?,?) ,XIC(PV_Security.Timers[7].DN) OTU(PV_Security.Bits.18) ];
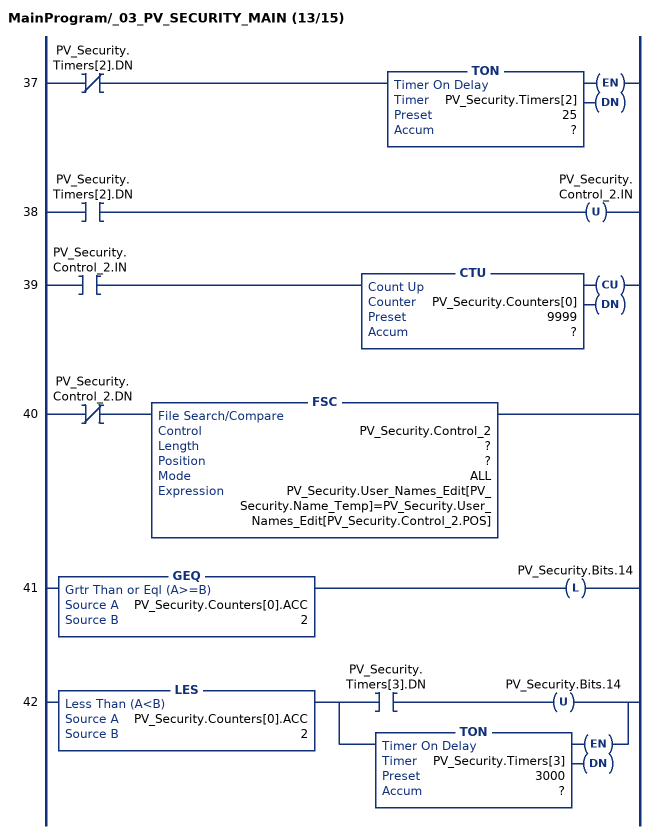
   37: XIO(PV_Security.Timers[2].DN)TON(PV_Security.Timers[2],?,?);
   38: XIC(PV_Security.Timers[2].DN)OTU(PV_Security.Control_2.IN);
   39: XIC(PV_Security.Control_2.IN)CTU(PV_Security.Counters[0],?,?);
   40: XIO(PV_Security.Control_2.DN)FSC(PV_Security.Control_2,?,?,ALL,PV_Security.User_Names_Edit[PV_Security.Name_Temp]=PV_Security.User_Names_Edit[PV_Security.Control_2.POS]);
   41: GEQ(PV_Security.Counters[0].ACC,2)OTL(PV_Security.Bits.14);
   42: LES(PV_Security.Counters[0].ACC,2)[XIC(PV_Security.Timers[3].DN) OTU(PV_Security.Bits.14) ,TON(PV_Security.Timers[3],?,?) ];
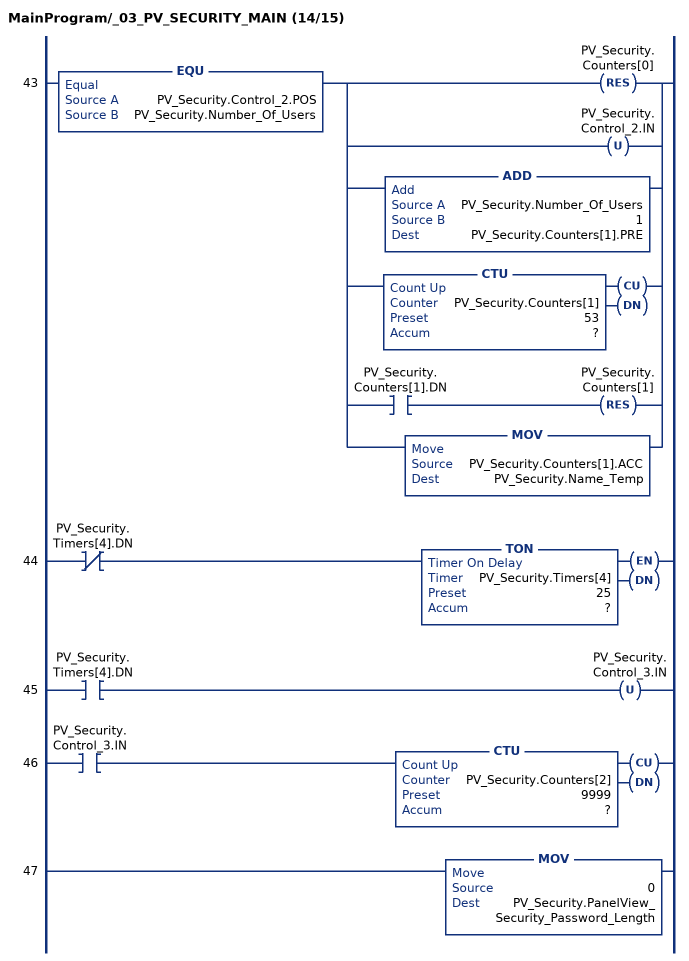
   43: EQU(PV_Security.Control_2.POS,PV_Security.Number_Of_Users)[RES(PV_Security.Counters[0]) ,OTU(PV_Security.Control_2.IN) ,ADD(PV_Security.Number_Of_Users,1,PV_Security.Counters[1].PRE) ,CTU(PV_Security.Counters[1],?,?) ,XIC(PV_Security.Counters[1].DN) RES(PV_Security.Counters[1]) ,MOV(PV_Security.Counters[1].ACC,PV_Security.Name_Temp) ];
   44: XIO(PV_Security.Timers[4].DN)TON(PV_Security.Timers[4],?,?);
   45: XIC(PV_Security.Timers[4].DN)OTU(PV_Security.Control_3.IN);
   46: XIC(PV_Security.Control_3.IN)CTU(PV_Security.Counters[2],?,?);
   47: MOV(0,PV_Security.PanelView_Security_Password_Length);
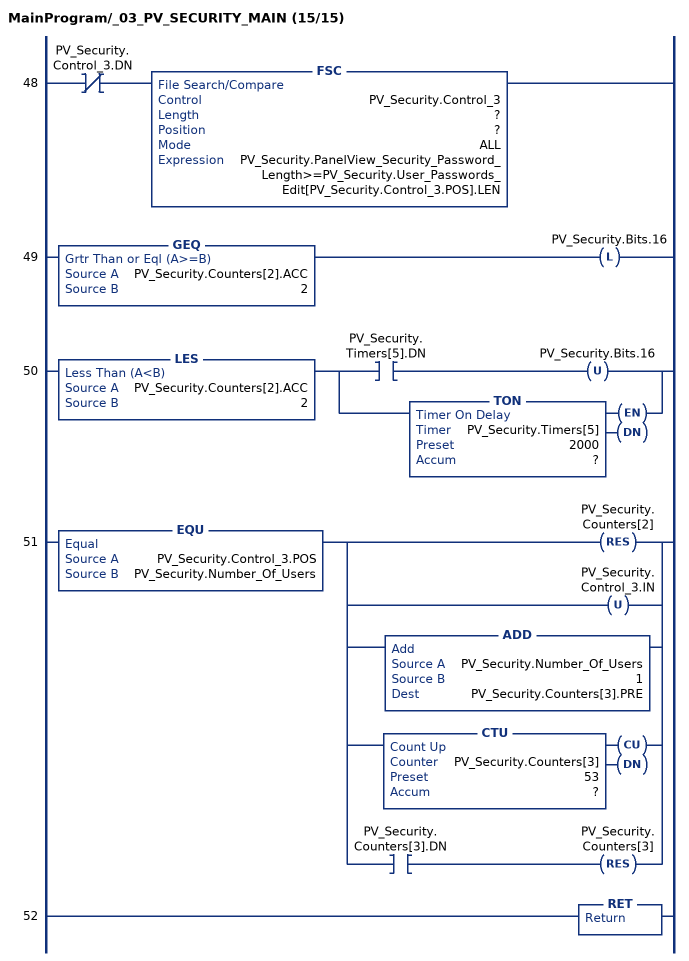
   48: XIO(PV_Security.Control_3.DN)FSC(PV_Security.Control_3,?,?,ALL,PV_Security.PanelView_Security_Password_Length>=PV_Security.User_Passwords_Edit[PV_Security.Control_3.POS].LEN);
   49: GEQ(PV_Security.Counters[2].ACC,2)OTL(PV_Security.Bits.16);
   50: LES(PV_Security.Counters[2].ACC,2)[XIC(PV_Security.Timers[5].DN) OTU(PV_Security.Bits.16) ,TON(PV_Security.Timers[5],?,?) ];
   51: EQU(PV_Security.Control_3.POS,PV_Security.Number_Of_Users)[RES(PV_Security.Counters[2]) ,OTU(PV_Security.Control_3.IN) ,ADD(PV_Security.Number_Of_Users,1,PV_Security.Counters[3].PRE) ,CTU(PV_Security.Counters[3],?,?) ,XIC(PV_Security.Counters[3].DN) RES(PV_Security.Counters[3]) ];
   52: RET();
END_ROUTINE
